(* IEC 61131-3 sources: daoli-st-library/DL_Process (part 58) *)

(* ---- FB_DL_VacuumBakeOutSeq.st ---- *)
(*
  组件名 Component   : FB_DL_VacuumBakeOutSeq
  子库 Sublibrary    : DL_Process
  版本 Version       : 1.0.0
  兼容性 Platform    : CODESYS 3.5 / TwinCAT 3 / 汇川 InoProShop / Machine Expert（仅 Standard.library）
  功能 Function      : 真空烘烤顺控（锂电/半导体共性，自研行业池）：
                       1) 升温相（eRampUp）：温度需求按 fRampRateKMin 斜率逼近
                       fSoakTempC，腔压 < fSoakPressMaxPa 才视为升温有效；
                       2) 保温保压相（eSoak）：温度需求保持 fSoakTempC，腔压超上限
                       持续 tPressDevTo → 故障锁存；保温计时到 → 进压升率判漏相；
                       3) 压升率判漏相（eRorMeas）：窗始取腔压快照，窗长 tRorWin 到
                       → 压升率 = (腔压 - 快照) / 窗长，超 fRorFailPaS → 故障（判漏
                       不合格）；不超 → 终点判据达成，进降温相；
                       4) 降温放气相（eCoolVent）：需求温度按斜率降至 fEndTempC 后
                       开放气阀驻留 tVentDur → eDone。
  边界 Boundary      : ① 本件只出温度需求/阀门指令，不写物理 IO，不内嵌温控回路；
                       ② 压升率除法前置域闸：tRorWin 秒值下限 0.1 s（常量护栏）；
                       ③ 各相计时独立 TON 实例（禁跨相复用）；压升率窗始快照在
                       进相首拍写定，锁存回放不重扫；
                       ④ 故障锁存解除唯一路径 = bReset 上升沿（输入引脚，恒可达）；
                       ⑤ 无全局变量引用、无外部变量声明、无物理地址寻址。
  依赖 Depends       : Standard.library（R_TRIG / TON）
  溯源 Origin        : 道莅自研 clean-room（自研行业池：锂电/半导体真空烘烤共性
                       语义，零外部代码行复制）
  码位 Code          : 16#06_0_BF（Process 段 0006，B 子带 BF 格）
  码表 Error codes（本件格 06_0_BF，单轨子道：故障 0x02BF / 信息 0x01BF）:
    16#0006_02BF 故障级：烘烤顺控故障总码（保压越限 / 压升率判漏不合格 /
                 组态非法 / 输入非有限），锁存至复位
    16#0006_01BF 信息级：压升率判漏通过沿（进降温相迁移拍）
  修订历史 Revision  :
    2026-11-19  v1.0.0  R44 首版（批次 4 · 序号 16）
*)

TYPE E_DL_VboPhase :
(
    eIdle     := 0,   // 空闲：未使能 / Idle, not enabled
    eRampUp   := 10,  // 升温：斜坡逼近保温温度 / Ramping to soak temperature
    eSoak     := 20,  // 保温保压：保持温度与压力 / Soaking temperature and pressure
    eRorMeas  := 30,  // 判漏：压升率测量窗 / Rate-of-rise measurement window
    eCoolVent := 40,  // 降温放气：斜坡降温 + 放气 / Cooling and venting
    eDone     := 50,  // 完成：终点驻留 / Done, endpoint held
    eFault    := 90   // 故障：总码锁存 / Fault, latched
);
END_TYPE

FUNCTION_BLOCK FB_DL_VacuumBakeOutSeq
VAR_INPUT
    bEnable      : BOOL;                   // 使能（电平）[-] / Enable
    bReset       : BOOL;                   // 上升沿清故障锁存 [-] / Reset edge
    fChamberTempC: REAL;                   // 腔体实测温度 [摄氏度] / Chamber temperature
    fChamberPressPa: REAL;                 // 腔体实测压力 [帕斯卡] / Chamber pressure
    fSoakTempC   : REAL := 80.0;           // 保温温度 [摄氏度] / Soak temperature
    fEndTempC    : REAL := 35.0;           // 降温终点温度 [摄氏度] / Cool-down end temperature
    fRampRateKMin: REAL := 2.0;            // 升降温斜率 [开尔文/分] / Ramp rate
    fSoakPressMaxPa: REAL := 50.0;         // 保温压力上限 [帕斯卡] / Soak pressure ceiling
    fRorFailPaS  : REAL := 5.0;            // 压升率判漏限 [帕/秒] / Rate-of-rise fail limit
    tSoakDur     : TIME := T#24H;          // 保温时长 [毫秒] / Soak duration
    tRorWin      : TIME := T#60S;          // 压升率测量窗 [毫秒] / ROR measurement window
    tPressDevTo  : TIME := T#30S;          // 保压越限确认窗 [毫秒] / Pressure deviation timeout
    tVentDur     : TIME := T#60S;          // 放气驻留 [毫秒] / Vent dwell
    tCycle       : TIME := T#1S;           // 扫描周期 [毫秒] / Scan cycle time
END_VAR
VAR_OUTPUT
    fTempDemandC : REAL;                   // 温度需求输出 [摄氏度] / Temperature demand
    bPumpCmd     : BOOL;                   // 抽真空维持指令（升温/保温/判漏相）[-] / Vacuum maintain command
    bVentCmd     : BOOL;                   // 放气阀指令（放气驻留相电平）[-] / Vent valve command
    fRorPaS      : REAL;                   // 实测压升率 [帕/秒] / Measured rate of rise
    ePhase       : E_DL_VboPhase;          // 相位出口，段尾单点映射 / Phase outlet
    bError       : BOOL;                   // 故障锁存标志 [-] / Fault latch flag
    uErrId       : UDINT;                  // 事件码，0 = 无事件 / Event code
END_VAR
VAR
    rtReset  : R_TRIG;                     // 复位沿实例，段 0 无条件刷新 / Reset edge
    tonSoakDur: TON;                       // 保温计时（独立实例） / Soak duration timer
    tonRorWin : TON;                       // 压升率测量窗（独立实例） / ROR window timer
    tonPressDevTo: TON;                    // 保压越限确认（专用超时件命名） / Pressure timeout
    tonVentDur: TON;                       // 放气驻留计时（独立实例） / Vent dwell timer
    _ePhase : E_DL_VboPhase := E_DL_VboPhase.eIdle;    // 内部相位（CASE 唯一写入目标）/ Internal phase
    _fPressSnap: REAL;                     // 判漏窗始压力快照 [帕斯卡] / Window-start pressure snapshot
    _fPressStart: REAL;                    // 保温起点压力快照 [帕斯卡] / Soak-start pressure snapshot
    _bFault : BOOL;                        // 故障锁存位（锁存量） / Latched fault bit
    _uFault : UDINT;                       // 故障码锁存（锁存量） / Latched fault code
    _bCfgBad: BOOL;                        // 组态非法当拍量 [-] / Config illegal flag
    _bNonFin: BOOL;                        // 输入非有限当拍量 [-] / Non-finite input flag
    _bSnapDone: BOOL;                      // 判漏快照已取标志 [-] / Snapshot taken flag
END_VAR
VAR CONSTANT
    DL_WIN_MIN_S : REAL := 0.1;            // 测量窗秒值下限 [秒] / Window seconds floor
    DL_SEC_PER_MIN: REAL := 60.0;          // 秒 → 分换算系数 [秒/分] / Seconds per minute
    DL_MS_PER_S  : REAL := 1000.0;         // 毫秒 → 秒换算系数 [毫秒/秒] / Milliseconds per second
    DL_ABS_MAX   : REAL := 1.0E30;         // 有限值判定上界 [工程单位] / Finite bound
    DL_ZERO      : REAL := 0.0;            // 零常量 [工程单位] / Zero constant
END_VAR

(* —— 段 0｜沿与定时器每拍无条件刷新（禁置于 IF/CASE 内；各相独立实例禁复用） —— *)
rtReset(CLK := bReset);
tonSoakDur   (IN := (_ePhase = E_DL_VboPhase.eSoak) AND (NOT _bFault), PT := tSoakDur);
tonRorWin    (IN := (_ePhase = E_DL_VboPhase.eRorMeas) AND (NOT _bFault), PT := tRorWin);
tonPressDevTo(IN := (_ePhase = E_DL_VboPhase.eSoak) AND (fChamberPressPa > fSoakPressMaxPa)
              AND (NOT _bFault), PT := tPressDevTo);
tonVentDur   (IN := (_ePhase = E_DL_VboPhase.eCoolVent) AND (NOT _bFault), PT := tVentDur);

(* —— 段 1｜瞬时量预清零（锁存量 _bFault/_uFault/fTempDemandC/_fPressSnap 不入清单） —— *)
uErrId   := 16#0000_0000;
_bCfgBad := FALSE;
_bNonFin := FALSE;

(* —— 段 2｜复位沿：故障一次性清干净，相位回空闲，阀门指令撤销 —— *)
IF rtReset.Q THEN
    _bFault := FALSE;
    _uFault := 16#0000_0000;
    bVentCmd := FALSE;
    bPumpCmd := FALSE;
    _ePhase := E_DL_VboPhase.eIdle;
END_IF

(* —— 段 3｜组态闸与非有限判据（覆盖全部参与判据换算引脚） —— *)
IF (fRampRateKMin <= DL_ZERO) OR (fRorFailPaS <= DL_ZERO) OR (tSoakDur = T#0S)
   OR (tRorWin = T#0S) OR (tPressDevTo = T#0S) OR (tVentDur = T#0S) OR (tCycle = T#0S)
   OR (fSoakTempC <= fEndTempC) THEN
    _bCfgBad := TRUE;
END_IF
IF (fChamberTempC <> fChamberTempC) OR ((fChamberTempC - fChamberTempC) <> DL_ZERO)
   OR (fChamberPressPa <> fChamberPressPa) OR ((fChamberPressPa - fChamberPressPa) <> DL_ZERO) THEN
    _bNonFin := TRUE;
END_IF

(* —— 段 4｜主状态机：七态全覆盖 + ELSE 兜底 —— *)
CASE _ePhase OF

E_DL_VboPhase.eIdle:
    fTempDemandC := fChamberTempC;       // 空闲相：需求跟随实测（不驱动）
    bPumpCmd := FALSE;
    bVentCmd := FALSE;
    IF bEnable AND (NOT _bCfgBad) THEN
        _bSnapDone := FALSE;
        fRorPaS := DL_ZERO;
        _ePhase := E_DL_VboPhase.eRampUp;
    ELSIF bEnable AND _bCfgBad THEN
        _bFault := TRUE;
        _uFault := 16#0006_02BF;
        bError  := TRUE;
        _ePhase := E_DL_VboPhase.eFault;
    END_IF

E_DL_VboPhase.eRampUp:
    bPumpCmd := TRUE;
    bVentCmd := FALSE;
    (* 温度需求斜率逼近：每拍步长 = 斜率 × 周期（分 → 秒换算，除子域闸已过） *)
    fTempDemandC := MIN(fTempDemandC + fRampRateKMin * (TIME_TO_REAL(tCycle) / DL_MS_PER_S)
                        / DL_SEC_PER_MIN, fSoakTempC);
    IF _bNonFin THEN
        _bFault := TRUE;
        _uFault := 16#0006_02BF;
        bError  := TRUE;
        _ePhase := E_DL_VboPhase.eFault;
    ELSIF NOT bEnable THEN
        _ePhase := E_DL_VboPhase.eIdle;  // 使能撤销回空闲
    ELSIF (fChamberTempC >= fSoakTempC) AND (fChamberPressPa <= fSoakPressMaxPa) THEN
        _fPressStart := fChamberPressPa; // 保温起点压力快照
        _ePhase := E_DL_VboPhase.eSoak;  // 迁出：温度达保温且压力已入保压域
    END_IF

E_DL_VboPhase.eSoak:
    bPumpCmd := TRUE;
    bVentCmd := FALSE;
    fTempDemandC := fSoakTempC;          // 保温相需求定值
    IF _bNonFin OR tonPressDevTo.Q THEN
        _bFault := TRUE;                 // 保压越限或输入非法：锁存
        _uFault := 16#0006_02BF;
        bError  := TRUE;
        _ePhase := E_DL_VboPhase.eFault;
    ELSIF NOT bEnable THEN
        _ePhase := E_DL_VboPhase.eIdle;  // 使能撤销回空闲
    ELSIF tonSoakDur.Q THEN
        _bSnapDone := FALSE;             // 保温时长到：进判漏相，快照待取
        _ePhase := E_DL_VboPhase.eRorMeas;
    END_IF

E_DL_VboPhase.eRorMeas:
    bPumpCmd := TRUE;
    bVentCmd := FALSE;
    fTempDemandC := fSoakTempC;
    IF _bNonFin THEN
        _bFault := TRUE;
        _uFault := 16#0006_02BF;
        bError  := TRUE;
        _ePhase := E_DL_VboPhase.eFault;
    ELSIF NOT _bSnapDone THEN
        _fPressSnap := fChamberPressPa;  // 窗始快照：进相首拍写定（锁存回放不重扫）
        _bSnapDone := TRUE;
    ELSIF tonRorWin.Q THEN
        (* 压升率 = (腔压 - 窗始快照) / 窗长秒值（除子 = 窗长，常量护栏下限已过） *)
        fRorPaS := (fChamberPressPa - _fPressSnap)
                   / MAX(TIME_TO_REAL(tRorWin) / DL_MS_PER_S, DL_WIN_MIN_S);
        IF fRorPaS > fRorFailPaS THEN
            _bFault := TRUE;             // 判漏不合格：锁存（禁按当下输入重推断）
            _uFault := 16#0006_02BF;
            bError  := TRUE;
            _ePhase := E_DL_VboPhase.eFault;
        ELSE
            uErrId := 16#0006_01BF;      // 信息级：判漏通过沿
            _ePhase := E_DL_VboPhase.eCoolVent;   // 终点判据达成：进降温放气
        END_IF
    END_IF

E_DL_VboPhase.eCoolVent:
    bPumpCmd := FALSE;
    (* 温度需求斜率下降，降至终点温度前放气阀不开（先降温后放气） *)
    IF fTempDemandC > fEndTempC THEN
        fTempDemandC := MAX(fTempDemandC - fRampRateKMin * (TIME_TO_REAL(tCycle) / DL_MS_PER_S)
                            / DL_SEC_PER_MIN, fEndTempC);
        bVentCmd := FALSE;
    ELSE
        bVentCmd := TRUE;                // 需求到终点温度：开放气阀驻留
    END_IF
    IF _bNonFin THEN
        _bFault := TRUE;
        _uFault := 16#0006_02BF;
        bError  := TRUE;
        _ePhase := E_DL_VboPhase.eFault;
    ELSIF bVentCmd AND tonVentDur.Q THEN
        _ePhase := E_DL_VboPhase.eDone;  // 迁出：放气驻留完成
    ELSIF NOT bEnable THEN
        _ePhase := E_DL_VboPhase.eIdle;  // 使能撤销回空闲
    END_IF

E_DL_VboPhase.eDone:
    bPumpCmd := FALSE;
    bVentCmd := FALSE;                   // 完成相：阀门指令全撤（安全侧）
    IF NOT bEnable THEN
        _ePhase := E_DL_VboPhase.eIdle;  // 使能撤销回空闲（待机可返回路径）
    END_IF

E_DL_VboPhase.eFault:
    bPumpCmd := FALSE;
    bVentCmd := FALSE;
    bError := TRUE;
    ;                                    // 故障相驻留：只认复位沿（段 2 迁出）

ELSE
    _bFault := TRUE;                     // 兜底：非法相位锁存
    _uFault := 16#0006_02BF;
    bError  := TRUE;
    _ePhase := E_DL_VboPhase.eFault;
END_CASE

(* —— 段 5｜相位出口单点映射 —— *)
ePhase := _ePhase;
END_FUNCTION_BLOCK

(* ---- FB_DL_VacuumChamberSeq.st ---- *)
(*==============================================================================
 * 组件名称 (Component)  : FB_DL_VacuumChamberSeq
 * 所属子库 (Sublibrary) : DL_Process
 * 前缀     (Prefix)     : FB_DL_
 * 当前版本 (Version)    : 1.0.0
 * 兼容性   (Platform)   : CODESYS 3.5 / TwinCAT 3 / 汇川 InoProShop / Schneider
 *                         Machine Expert；纯 IEC 61131-3（第 3 版），
 *                         仅依赖标准库 TON / R_TRIG / ABS，零厂商方言
 * 作者     (Author)     : 道莅代码库 · PLC编程专家（R31）
 * 开源溯源 (Origin)     : 真空腔体抽真空顺控公开工艺语义（行业池），
 *                         道莅 clean-room 防御性实现，未复制任何外部源码行
 * 功能描述 (Function)   : 纯真空腔体五相顺控原子（不含工艺加热）：粗抽至
 *                         粗抽阈值 → 精抽至目标（迟滞防边界抖动）→ 检漏
 *                         （消费 bLeakOk）→ 放气（数字阀经缓启时序等价
 *                         斜坡限幅防冲击）→ 完成。相转换本拍复验数据源
 *                         （R42）；步超时锁故障；中止安全次序写死：
 *                         先停泵、延时后才开放气阀。
 * 组合建议 (Composition): 与库内 FB_DL_SlitValveInterlock 组合使用——本件
 *                         给出真空工艺时序，闸阀联锁由该件承担，二者经
 *                         bLeakOk/泵指令引脚对接，不互相内嵌。
 * 状态机   (States)     : eIdle/eRough/eFine/eLeakTest/eVent/eFault，
 *                         CASE 带 ELSE 锁安全侧（全阀关、全泵停）。
 * 码位     (Codes)      : 16#0005_009E 信息级：压强数据非有限冻结当前相、
 *                                      迟滞等待提示（不置 bError）
 *                         16#0005_009F 故障级：相超时
 *                         16#0005_00A0 故障级：联锁违例（非空闲相重启）
 *                         16#0005_00A1 故障级：状态非法（ELSE 兜底，锁存）
 *                         16#0005_00A2 保留未启用（码表与实现对齐）
 * 边界防错 (Boundary)   : 1 压强非有限（x<>x 自反判加幅值界）冻结当前相；
 *                         2 精抽到位判定带迟滞：超回差即回信息级等待；
 *                         3 TON/R_TRIG 实例每拍无条件刷新，按相断输入；
 *                         4 CASE 带 ELSE 锁安全侧；
 *                         5 故障锁存可达解除路径：中止沿复归待机；
 *                         6 相转换本拍复验数据源（R42）。
 * 修订历史 (Revision)   : 2026-11-18 v1.0.0 首版入库（R31 · 阶段三 · 序 12）
 *==============================================================================*)

(*------------------------------------------------------------------------------
 * 枚举: E_DL_VacPhase（归属本功能块，同文件发布，全库唯一属主）
 *----------------------------------------------------------------------------*)
TYPE E_DL_VacPhase :
(
    eIdle     := 0,    // 空闲：全泵停全阀关 / Idle, all pumps and valves off
    eRough    := 10,   // 粗抽相：粗抽泵运行 / Rough phase, rough pump running
    eFine     := 20,   // 精抽相：精抽泵运行 / Fine phase, fine pump running
    eLeakTest := 30,   // 检漏相：泵停隔离等待结论 / Leak test, pumps off, isolated
    eVent     := 40,   // 放气相：缓启时序后开阀 / Vent phase, valve after ramp delay
    eFault    := 99    // 故障：锁定等待中止复位 / Fault, latched until abort reset
);
END_TYPE

(*==============================================================================
 * 功能块: FB_DL_VacuumChamberSeq
 * 调用约定: 每个扫描周期无条件调用一次；压强信号经引脚注入。
 *==============================================================================*)
FUNCTION_BLOCK FB_DL_VacuumChamberSeq
VAR_INPUT
    bStart   : BOOL := FALSE;         // 启动沿（空闲相受理）/ Start edge, accepted in idle
    bAbort   : BOOL := FALSE;         // 中止沿：任意相安全退出 / Abort edge, safe exit from any phase
    fPNow    : REAL := 101325.0;      // 腔体当前压强 [帕] / Chamber current pressure [Pa]
    fPTgt    : REAL := 10.0;          // 精抽目标压强 [帕] / Fine target pressure [Pa]
    fPRough  : REAL := 500.0;         // 粗抽切换阈值 [帕] / Rough crossover threshold [Pa]
    bLeakOk  : BOOL := FALSE;         // 检漏结论注入（外部检漏件）/ Leak verdict injected by caller
    tStepMax : TIME := T#600S;        // 单相超时 [毫秒] / Per-phase timeout [ms]
    tVentRamp: TIME := T#5S;          // 放气缓启时序 [毫秒]（斜坡限幅等价实现）/ Vent ramp delay [ms]
END_VAR
VAR_OUTPUT
    ePhase    : E_DL_VacPhase;        // 当前相状态 / Current phase
    bPumpRough: BOOL;                 // 粗抽泵指令 / Rough pump command
    bPumpFine : BOOL;                 // 精抽泵指令 / Fine pump command
    bVent     : BOOL;                 // 放气阀指令 / Vent valve command
    bDone     : BOOL;                 // 流程完成单拍脉冲（R27）/ Sequence done one-scan pulse
    bError    : BOOL;                 // 故障标志，与故障级码配对（R45）/ Fault flag paired with fault codes
    uErrorId  : UDINT;                // 错误码，0 = 无错 / Error code, 0 = none
END_VAR
VAR
    rTrigStart: R_TRIG;               // 启动沿检测，每拍无条件刷新 / Start edge detector, refreshed every scan
    rTrigAbort: R_TRIG;               // 中止沿检测，每拍无条件刷新 / Abort edge detector, refreshed every scan
    tonPhase  : TON;                  // 相超时定时器，每拍无条件刷新 / Phase timeout timer, refreshed every scan
    tonVent   : TON;                  // 放气缓启定时器，每拍无条件刷新 / Vent ramp timer, refreshed every scan
    eStatePrev: E_DL_VacPhase;        // 上一拍相快照 / Previous phase snapshot
    bStepRst  : BOOL;                 // 相切换拍单拍断超时输入 / One-scan timeout break on phase change
    bDataOk   : BOOL;                 // 压强三点有效性 / Three pressure points validity
    bHystWait : BOOL;                 // 迟滞等待标志 / Hysteresis waiting flag
    bAborted  : BOOL;                 // 中止退出路径标志 / Abort exit path flag
    uCodeLatch: UDINT;                // 故障级锁存码 / Latched fault code
    bInit     : BOOL := TRUE;         // 首扫标志 / First-scan flag
END_VAR
VAR CONSTANT
    DL_VCS_FIN    : REAL := 1.0E30;   // REAL 有限幅值判界 / REAL finiteness magnitude bound
    DL_VCS_HYST   : REAL := 1.1;      // 精抽迟滞回差系数（超回差回等待）/ Fine hysteresis back factor
    DL_VCS_PATM   : REAL := 90000.0;  // 放气完成压强阈 [帕] / Vent complete pressure threshold [Pa]
END_VAR

// ---- 段 1｜边沿与定时器实例无条件周期刷新（红线：禁入条件分支）----------------
rTrigStart(CLK := bStart);                            // 启动沿检测 / Start edge detection
rTrigAbort(CLK := bAbort);                            // 中止沿检测 / Abort edge detection
tonVent(IN := (ePhase = eVent), PT := tVentRamp);     // 缓启计时按相断输入 / Ramp timing input per phase
tonPhase(IN := (ePhase <> eIdle) AND (ePhase <> eFault) AND (ePhase <> eVent)
         AND (NOT bStepRst), PT := tStepMax);         // 相超时计时，相切换拍断输入 / Phase timeout timing

// ---- 段 2｜相切换检测与数据有效性 ----------------------------------------------
bStepRst := (ePhase <> eStatePrev) OR bInit;          // 相变化即断输入 / Phase change breaks timing input
eStatePrev := ePhase;                                 // 快照留痕 / Snapshot previous phase
bInit := FALSE;                                       // 清首扫标志 / Clear first-scan flag
bDataOk := (fPNow = fPNow) AND (fPTgt = fPTgt) AND (fPRough = fPRough)
       AND (ABS(fPNow) < DL_VCS_FIN) AND (ABS(fPTgt) < DL_VCS_FIN)
       AND (ABS(fPRough) < DL_VCS_FIN);               // 压强三点有限 / Three points finite

// ---- 段 3｜中止沿统一入口：先停泵、缓启延时后才放气（安全次序写死）--------------
IF rTrigAbort.Q AND (ePhase <> eIdle) THEN
    ePhase   := eVent;                                // 转放气相执行退出 / To vent phase for exit
    bAborted := TRUE;                                 // 登记中止路径 / Mark abort path
END_IF

// ---- 段 4｜状态机（CASE 带 ELSE 锁安全侧：全泵停全阀关）--------------------------
CASE ePhase OF
    eIdle:
        bPumpRough := FALSE;                          // 空闲全停 / All off in idle
        bPumpFine  := FALSE;                          // 空闲全停 / All off in idle
        bVent      := FALSE;                          // 空闲阀关 / Valve closed in idle
        bDone      := FALSE;                          // 清完成脉冲 / Clear done pulse
        bAborted   := FALSE;                          // 清中止标志 / Clear abort flag
        IF rTrigStart.Q AND bDataOk AND (fPTgt < fPRough) THEN
            ePhase := eRough;                         // 数据合法且目标低于切换阈才启动 / Legal data and sane targets
        END_IF
    eRough:
        bPumpRough := bDataOk AND NOT bAborted;       // 粗抽泵指令带数据门控 / Rough pump gated by data
        bPumpFine  := FALSE;                          // 精抽泵停 / Fine pump off
        bVent      := FALSE;                          // 阀关 / Valve closed
        IF NOT bDataOk THEN
            uErrorId := 16#0005_009E;                 // 信息级：数据非有限冻结当前相 / Info: non-finite freezes phase
        ELSIF tonPhase.Q THEN
            ePhase := eFault;                         // 相超时锁故障 / Phase timeout, fault
            uCodeLatch := 16#0005_009F;               // 码位：相超时 / Code: phase timeout
        ELSIF bDataOk AND (fPNow <= fPRough) THEN
            ePhase := eFine;                          // 复验后转精抽（R42）/ Recheck then to fine
        END_IF
    eFine:
        bPumpRough := FALSE;                          // 粗抽泵停（交叉点切换）/ Rough pump off at crossover
        bPumpFine  := bDataOk AND NOT bAborted;       // 精抽泵指令带数据门控 / Fine pump gated by data
        bVent      := FALSE;                          // 阀关 / Valve closed
        bHystWait  := bDataOk AND (fPNow > fPTgt * DL_VCS_HYST); // 超回差等待 / Beyond hysteresis, wait
        IF NOT bDataOk THEN
            uErrorId := 16#0005_009E;                 // 信息级：数据非有限冻结当前相 / Info: non-finite freezes phase
        ELSIF tonPhase.Q THEN
            ePhase := eFault;                         // 相超时锁故障 / Phase timeout, fault
            uCodeLatch := 16#0005_009F;               // 码位：相超时 / Code: phase timeout
        ELSIF bHystWait THEN
            uErrorId := 16#0005_009E;                 // 信息级：迟滞等待提示 / Info: hysteresis waiting
        ELSIF bDataOk AND (fPNow <= fPTgt) THEN
            ePhase := eLeakTest;                      // 复验后转检漏（R42）/ Recheck then to leak test
        END_IF
    eLeakTest:
        bPumpRough := FALSE;                          // 检漏隔离全泵停 / Isolated, all pumps off
        bPumpFine  := FALSE;                          // 检漏隔离全泵停 / Isolated, all pumps off
        bVent      := FALSE;                          // 阀关 / Valve closed
        IF tonPhase.Q THEN
            ePhase := eFault;                         // 相超时锁故障 / Phase timeout, fault
            uCodeLatch := 16#0005_009F;               // 码位：相超时 / Code: phase timeout
        ELSIF bLeakOk THEN
            ePhase := eVent;                          // 检漏合格转放气 / Leak OK, to vent
        END_IF
    eVent:
        bPumpRough := FALSE;                          // 放气相全泵停 / All pumps off in vent
        bPumpFine  := FALSE;                          // 放气相全泵停 / All pumps off in vent
        bVent      := tonVent.Q;                      // 缓启时序满才开阀（先停泵后放气）/ Valve after ramp, pumps first
        IF (NOT bAborted) AND bDataOk AND (fPNow >= DL_VCS_PATM) THEN
            ePhase := eIdle;                          // 正常放气完成回待机 / Normal vent complete
            bDone := TRUE;                            // 完成单拍脉冲 / One-scan done pulse
        ELSIF bAborted AND tonVent.Q THEN
            ePhase := eIdle;                          // 中止退出回待机 / Abort exit back to idle
            bDone := FALSE;                           // 中止不置完成 / Abort never sets done
        END_IF
    eFault:
        bPumpRough := FALSE;                          // 故障安全侧全停 / Fault safe side all off
        bPumpFine  := FALSE;                          // 故障安全侧全停 / Fault safe side all off
        bVent      := FALSE;                          // 故障安全侧阀关 / Fault safe side valve closed
        bDone      := FALSE;                          // 故障清完成 / Fault clears done
        IF rTrigAbort.Q THEN
            ePhase := eIdle;                          // 可达解除路径：中止沿复归 / Reachable release: abort edge
            uCodeLatch := 16#0000_0000;               // 清锁存码 / Clear latched code
        END_IF
    ELSE
        ePhase := eFault;                             // 非法状态兜底 / Illegal state fallback
        uCodeLatch := 16#0005_00A1;                   // 码位：状态非法 / Code: illegal state
END_CASE

// ---- 段 5｜联锁违例防御：非空闲相受理启动沿 --------------------------------------
IF rTrigStart.Q AND (eStatePrev <> eIdle) AND (ePhase <> eIdle) AND (ePhase <> eFault) THEN
    ePhase := eFault;                                 // 违例锁故障 / Violation latches fault
    uCodeLatch := 16#0005_00A0;                       // 码位：联锁违例 / Code: interlock violation
END_IF

// ---- 段 6｜错误码装配：故障锁存回放优先，信息级居次 ------------------------------
IF ePhase = eFault THEN
    bError   := TRUE;                                 // 故障标志配对（R45）/ Fault flag paired
    uErrorId := uCodeLatch;                           // 故障码锁存回放 / Latched fault code replayed
ELSIF (NOT bDataOk) OR bHystWait THEN
    bError   := FALSE;                                // 信息级不置故障 / Info never sets fault
    uErrorId := 16#0005_009E;                         // 信息级：冻结/迟滞等待 / Info: frozen or hysteresis wait
ELSE
    bError   := FALSE;                                // 无错清标志 / Clear fault flag
    uErrorId := 16#0000_0000;                         // 无码 / No code
END_IF
END_FUNCTION_BLOCK

(* ---- FB_DL_VavCouplingFeedforward.st ---- *)
(*==============================================================================
 * 组件名称 (Component)  : FB_DL_VavCouplingFeedforward
 * 所属子库 (Sublibrary) : DL_Process
 * 归属目录 (Directory)  : C:\Library\DL_Process
 * 当前版本 (Version)    : 1.0.0
 * 分类/来源标签         : 功能块（FUNCTION_BLOCK）· 暖通前馈 · 变风量耦合
 *                         industry-pool / hvac / vav / feedforward
 * 兼容性   (Platform)   : CODESYS 3.5 / TwinCAT 3 / 汇川 InoProShop / 施耐德
 *                         Machine Expert；仅用 Standard.library 的 ABS
 * 溯源声明 (Provenance) : 道莅自研 clean-room——只借公开规范条款与工程惯例，零代码行复制。
 * 功能一句话 (Summary)  : 送风温度偏离设计值时按显热守恒比例前馈修正风量
 *                         给定，替代反馈环慢慢追赶，防送风温度-风量耦合振荡。
 *
 * 功能描述 (Function)   : 显热守恒：风量与（室温设定 − 送风温度）成反比，
 *                         前馈量 = 设计风量 × 设计温差 ÷ 当前温差；当前温差
 *                         绝对值小于容差时视为近设计工况，恒等输出设计风量
 *                         并报信息级；输入非有限冻结输出（故障级）；送风
 *                         过热（温差反号）按最小风量保守输出；结果钳位到
 *                         风量上下限并报钳位码。内部状态与输出模式分离，
 *                         输出预置不触碰状态驻留量（R19）。
 * 与既有件边界 (Boundary): 本件只做静态前馈，不含反馈环与执行器控制；
 *                         VAV 盒反馈控制归 FB_DL_VavBoxCtrl，二者级联使用。
 * 码位说明 (Codes)      : 信息 16#0006_300A 近设计工况恒等输出设计风量
 *                         故障 16#0006_300B 输入非有限，输出冻结
 *                         故障 16#0006_300C 送风过热（温差反号），按最小风量保守
 *                         故障 16#0006_300D 结果越限已钳位到风量上下限
 *                         段 16#06_0_0A~0E 首槽信息级、次槽起故障级。
 * 依赖说明 (Depends)    : 无 DL_ 内部依赖；仅 Standard.library 的 ABS。
 * 红线自检 (Redline)    : 零全局依赖 ｜ 零 VAR_EXTERNAL ｜ 零 %I/%Q ｜ 纯 IEC 标准库
 *                         除法前强制判零（温差容差闸）｜ 浮点比较带 fEps 容差
 *                         NaN/Inf 精确判据拦截 ｜ ENUM 配 CASE 且 ELSE 兜底
 *                         全变量双语同行注释 ｜ 无定时器实例
 * 修订历史 (Revision)   : 2026-11-18  v1.0.0  首版入库（R32 · 批 3）
 *============================================================================*)

FUNCTION_BLOCK FB_DL_VavCouplingFeedforward
VAR_INPUT
    bRun        : BOOL;                     // 前馈使能，假则输出设计风量并停算 / Enable, FALSE outputs the design flow
    fTsaC       : LREAL;                    // 送风温度 [degC] / Supply air temperature
    fTsaDesignC : LREAL := 13.0;            // 设计送风温度 [degC] / Design supply air temperature
    fRoomSetC   : LREAL := 24.0;            // 室温设定 [degC] / Room setpoint
    fQDesign    : LREAL := 500.0;           // 设计风量 [m3/h] / Design airflow
    fQMin       : LREAL := 100.0;           // 最小风量 [m3/h] / Minimum airflow
    fQMax       : LREAL := 1200.0;          // 最大风量 [m3/h] / Maximum airflow
    fDtEps      : LREAL := 0.5;             // 温差容差 [K]，低于此视为近设计 / Delta-T tolerance
    fEps        : LREAL := 1.0E-6;          // 浮点判零容差 [实数域] / Floating zero tolerance
END_VAR
VAR_OUTPUT
    eMode   : (eBypass := 0, eAuto := 1);       // 模式枚举输出：旁路/自动 / Mode output enum
    fQFf    : LREAL;                    // 前馈风量给定 [m3/h] / Feedforward airflow setpoint
    bClamp  : BOOL;                     // 钳位标志，结果被上下限裁剪时为真 / TRUE when the result was clamped
    bValid  : BOOL;                     // 前馈有效标志，冻结期间为假 / TRUE when the output is valid
    bError  : BOOL;                     // 故障标志，与故障码配对 / Fault flag paired with codes
    uErrorId: UDINT;                    // 事件码，0 表示无事件 / Event code, zero means none
END_VAR
VAR
    _eState   : (eStBypass := 0, eStAuto := 1);     // 内部状态机：旁路/自动，输出预置不触碰 / Internal state, never pre-set
    fDtDesign : LREAL;  // 设计温差 [K]，室温设定减设计送风温度 / Design delta-T
    fDtNow    : LREAL;  // 当前温差 [K] / Current delta-T
    fRatio    : LREAL;  // 温差比 [比值]，设计温差除当前温差 / Delta-T ratio
    fQCalc    : LREAL;  // 计算风量 [m3/h] / Calculated airflow
    bSigOk    : BOOL;   // 输入有效标志 / Input validity flag
    uCode     : UDINT;  // 码位暂存，出口单点写入 [码] / Code staging
END_VAR

(* 段 1｜输出预置（不触碰 _eState 状态驻留量，R19 预清零清单纪律）/ Pre-set outputs, the state stays resident *)
fQFf    := fQDesign;                // 默认输出设计风量 / Default output is the design flow
bClamp  := FALSE;
bValid  := FALSE;
bError  := FALSE;
uErrorId := 16#0000_0000;
uCode   := 16#0000_0000;
eMode   := eBypass;                 // 模式输出随内部状态在出口刷新 / Mode output refreshed at the exit

(* 段 2｜温差导出与输入有效性（NaN 自反、Inf 上限、风量域正）/ Delta-T and validity *)
fDtDesign := fRoomSetC - fTsaDesignC;   // 设计温差导出 / Design delta-T
fDtNow    := fRoomSetC - fTsaC;         // 当前温差导出 / Current delta-T
bSigOk := (fTsaC = fTsaC) AND (fQDesign = fQDesign)             // NaN 自反判据 / NaN reflexivity
          AND (ABS(fTsaC) < 1.0E308) AND (ABS(fQDesign) < 1.0E308)   // Inf 上限判据 / Inf limit
          AND (fQDesign > fEps) AND (fQMin > 0.0) AND (fQMax > fQMin);   // 风量域约束 / Flow domain

(* 段 3｜状态机主分派（ENUM 配 CASE，ELSE 兜底）/ State dispatch with ELSE interception *)
CASE _eState OF

    eStBypass:
        (* 本拍行为：旁路保持设计风量；使能且数据有效拍 N+1 进自动 / Hold design flow; arm when enabled *)
        IF bRun AND bSigOk THEN
            _eState := eStAuto;         // 拍 N 旁路相满足条件，拍 N+1 转自动 / To auto next scan
        END_IF

    eStAuto:
        (* 本拍行为：按显热守恒算前馈；撤使能回旁路，数据无效冻结输出 / Compute feedforward; freeze on bad data *)
        IF NOT bRun THEN
            _eState := eStBypass;       // 拍 N+1 回旁路 / Back to bypass next scan
            fQFf := fQDesign;           // 旁路输出设计风量 / Bypass outputs design flow
        ELSIF NOT bSigOk THEN
            fQFf := fQDesign;           // 冻结：保持设计风量，不发异常值 / Freeze at design flow
            bValid := FALSE;            // 有效标志撤 / Withdraw validity
            uCode := 16#0006_300B;      // 故障级：输入非有限 / Fault: non-finite input
        ELSIF fDtNow < -fDtEps THEN
            fQFf := fQMin;              // 送风过热：保守最小风量 / Overheated supply: conservative minimum
            bValid := TRUE;
            uCode := 16#0006_300C;      // 故障级：温差反号 / Fault: reversed delta-T
        ELSE
            IF ABS(fDtNow) < fDtEps THEN
                fQFf := fQDesign;       // 近设计工况：恒等输出 / Near design: identity output
                bValid := TRUE;
                uCode := 16#0006_300A;  // 信息级：近设计恒等 / Info: near-design identity
            ELSE
                (* 除零前置闸：温差已过容差闸，此处防御复检再除 / Defensive recheck before the division *)
                IF ABS(fDtNow) > fEps THEN
                    fRatio := fDtDesign / fDtNow;   // 温差比 / Delta-T ratio
                    fQCalc := fQDesign * fRatio;    // 前馈风量 / Feedforward flow
                    IF fQCalc < fQMin THEN
                        fQCalc := fQMin;            // 钳下限 / Clamp to minimum
                        bClamp := TRUE;
                    ELSIF fQCalc > fQMax THEN
                        fQCalc := fQMax;            // 钳上限 / Clamp to maximum
                        bClamp := TRUE;
                    END_IF
                    fQFf := fQCalc;     // 前馈输出 / Feedforward output
                    bValid := TRUE;
                    IF bClamp THEN
                        uCode := 16#0006_300D;      // 故障级：结果已钳位 / Fault: clamped
                    END_IF
                ELSE
                    fQFf := fQMax;      // 防御路：温差趋零按最大风量 / Defensive: max flow as delta-T vanishes
                    bValid := TRUE;
                    uCode := 16#0006_300D;
                END_IF
            END_IF
        END_IF

ELSE
    _eState := eStBypass;               // 非法状态拦截回旁路 / Illegal state to bypass
    fQFf := fQDesign;                   // 保守输出设计风量 / Conservative design flow
    uCode := 16#0006_300B;              // 故障级：状态越界 / Fault: state out of range
END_CASE

(* 段 4｜出口装配 / Exit assembly *)
eMode := eBypass;                       // 出口刷新模式输出 / Refresh the mode output at the exit
IF _eState = eStAuto THEN
    eMode := eAuto;                     // 自动相映射 / Auto mapping
END_IF
bError := (uCode >= 16#0006_300B) AND (uCode <= 16#0006_300D);  // 故障级码段判定 / Fault band check
uErrorId := uCode;                      // 码位单点写入 / Single write point
END_FUNCTION_BLOCK

(* ---- FB_DL_VavDischargeAirReset.st ---- *)
(*
  FB_DL_VavDischargeAirReset  —  送风温度重置（末端阀位加权平均 → 送风设定值） / VAV discharge-air reset from terminal damper weighted mean
  分类 Category : DL_Process
  版本 Version  : 1.0.0
  来源 Source   : t1-2-oscat — 末端重置族零检索深化
  溯源 Origin   : clean-room 实现，未复制任何源码行
  功能 Function : 1) 末端阀位有效性门控：权重 = 有效末端数量（阀位域 [0,100] 且有限），
                  加权平均 fWMean := SUM(有效阀位)/有效末端数；
                  2) 重置律：fAirSet := fBaseSet + fResetSpan × fWMean/100，输出钳位
                  [fSetMin, fSetMax]，钳位发生置信息级 0494；
                  3) 权重和 = 0（全部末端无效）→ 防除零退回默认设定值 fBaseSet +
                  信息级 0492（不置故障）；
                  4) 部分末端无效置信息级 0493；非有限阀位 → 036B 锁存；
                  质量判定 CASE 全覆盖 + ELSE 兜底落 036C。
  边界 Boundary : ① 组态闸：uTermCnt < 1 或 > 8、fResetSpan < 0、设定钳位域颠倒 → 036A；
                  ② 除零防御：有效末端数 >= 1 过闸后才做除法；
                  ③ 无 GVL 依赖：纯引脚输入输出，无外部变量引用，无物理 IO 地址。
  依赖 Depends  : 仅 Standard.library（ABS / LREAL 算术）
  码表 Error codes（Process 段 0005，窗口 036A~036C / 0492~0494）:
    16#0005_036A 故障级：组态非法（末端数界外 / 重置幅值为负 / 钳位域颠倒），锁存至 bReset
    16#0005_036B 故障级：阀位非有限（NaN 自反判），锁存至 bReset
    16#0005_036C 故障级：质量判定落 ELSE 兜底（非法质量 ID），锁存至 bReset
    16#0005_0492 信息级：全部末端无效，退回默认设定值
    16#0005_0493 信息级：部分末端无效提示（有效末端照常聚合）
    16#0005_0494 信息级：设定值钳位提示
  修订历史 Revision :
    2026-11-19  v1.0.0  R41 首版（批次 4 · 序号 4）
*)

TYPE E_DL_VarResetQual :
(
    eAllValid   := 0,    // 全部末端有效 / All terminals valid
    ePartValid  := 10,   // 部分末端无效 / Some terminals invalid
    eNoneValid  := 20    // 全部末端无效 / No terminal valid
);
END_TYPE

FUNCTION_BLOCK FB_DL_VavDischargeAirReset
VAR_INPUT
    aDamper      : ARRAY[1..8] OF LREAL;  // 末端阀位 [0..100 %] / Terminal damper positions
    uTermCnt     : UINT := 1;         // 末端数 [个]，域 1..8 / Terminal count
    fBaseSet     : LREAL := 18.0;     // 基础送风设定 [°C] / Base discharge-air setpoint
    fResetSpan   : LREAL := 2.0;      // 重置幅值 [K]，域 >= 0（阀位 100% 时加满）/ Reset span
    fSetMin      : LREAL := 12.0;     // 设定值下限 [°C] / Setpoint lower clamp
    fSetMax      : LREAL := 26.0;     // 设定值上限 [°C] / Setpoint upper clamp
    bEnable      : BOOL := FALSE;     // 使能 [-] / Enable
    bReset       : BOOL := FALSE;     // 复位，上升沿清故障锁存 / Reset edge clears fault latch
END_VAR
VAR_OUTPUT
    fAirSet      : LREAL;             // 送风设定值出口 [°C] / Discharge-air setpoint outlet
    fWMean       : LREAL;             // 阀位加权平均 [0..100 %] / Weighted damper mean
    bValid       : BOOL;              // 输出有效标志 / Output valid flag
    bError       : BOOL;              // 故障锁存标志 / Fault latch flag
    nErrId       : UDINT;             // 事件码，0 = 无事件 / Event code
END_VAR
VAR
    rtReset      : R_TRIG;            // 复位沿实例，无条件刷新 / Reset edge instance
    _nCap        : INT;               // 生效末端数 [个] / Effective terminal count
    _nValid      : INT;               // 有效末端数 [个] / Valid terminal count
    _fSum        : LREAL;             // 阀位累加器 [0..100 %] / Damper sum accumulator
    _eQual       : E_DL_VarResetQual; // 质量判定（CASE 唯一写入目标）/ Quality verdict
    _bFault      : BOOL;              // 故障锁存位（锁存量）/ Latched fault bit
    _uFault      : UDINT;             // 故障码锁存（锁存量）/ Latched fault code
    _uInfo       : UDINT;             // 信息码，每拍重算 / Transient info code
    i            : INT;               // 聚合循环游标 [索引] / Aggregation loop cursor
    _nGuard      : INT;               // 聚合守卫计数 [次] / Aggregation guard counter
END_VAR

(* —— 段 0：沿实例无条件周期刷新（禁置于 IF/CASE 内） —— *)
rtReset(CLK := bReset);             // 复位沿（每拍必调）

(* —— 段 1：单拍量预清零（锁存量 _bFault/_uFault 不入清单，禁同拍抹除） —— *)
_uInfo := 16#0000_0000;             // 信息码每拍重算
bValid := FALSE;                    // 有效出口缺省 FALSE
nErrId := 16#0000_0000;             // 事件码缺省无事件
fAirSet := fBaseSet;                // 设定值缺省 = 默认设定值（退回口径）
fWMean := 0.0;                      // 均值缺省 0
_nValid := 0;                       // 有效计数清零
_fSum := 0.0;                       // 累加器清零
_nGuard := 0;                       // 守卫清零

(* —— 段 2：复位沿 + 组态域闸（当拍量判据） —— *)
IF rtReset.Q THEN                   // rtReset.Q = 当拍量
    _bFault := FALSE;               // 清故障锁存位
    _uFault := 16#0000_0000;        // 清故障锁存码
END_IF
_nCap := UINT_TO_INT(uTermCnt);     // 末端数快照
IF (_nCap < 1) OR (_nCap > 8) OR (fResetSpan < 0.0) OR (fSetMin >= fSetMax) THEN
    _uFault := 16#0005_036A;        // 故障级：组态非法
    _bFault := TRUE;
END_IF

(* —— 段 3：末端聚合（有效性门控；非有限 → 036B 锁存；守卫循环） —— *)
IF (NOT _bFault) AND (_nCap >= 1) AND (_nCap <= 8) THEN
    FOR i := 1 TO _nCap DO
        _nGuard := _nGuard + 1;     // 守卫递增
        IF _nGuard > 8 THEN
            EXIT;                   // 守卫兜底退出（理论不可达）
        END_IF
        IF (aDamper[i] <> aDamper[i]) OR ((aDamper[i] - aDamper[i]) <> (aDamper[i] - aDamper[i])) THEN
            _uFault := 16#0005_036B;    // 故障级：阀位非有限
            _bFault := TRUE;
        ELSIF (aDamper[i] >= 0.0) AND (aDamper[i] <= 100.0) THEN
            _nValid := _nValid + 1;     // 有效末端计数（权重 = 有效性门控）
            _fSum := _fSum + aDamper[i];    // 阀位累加
        END_IF
    END_FOR
END_IF

(* —— 段 4：质量判定（CASE 全覆盖 + ELSE 兜底） —— *)
IF (NOT _bFault) AND (_nCap >= 1) AND (_nCap <= 8) THEN
    IF _nValid = _nCap THEN
        _eQual := E_DL_VarResetQual.eAllValid;      // 全部有效
    ELSIF _nValid >= 1 THEN
        _eQual := E_DL_VarResetQual.ePartValid;     // 部分有效
        _uInfo := 16#0005_0493;                     // 信息级：部分无效提示
    ELSE
        _eQual := E_DL_VarResetQual.eNoneValid;     // 全部无效
    END_IF

    CASE _eQual OF
    E_DL_VarResetQual.eAllValid:
        fWMean := _fSum / INT_TO_LREAL(_nValid);    // 加权平均（分母 = 末端数 >= 1，防除零）
    E_DL_VarResetQual.ePartValid:
        fWMean := _fSum / INT_TO_LREAL(_nValid);    // 有效末端口径平均（同上防除零）
    E_DL_VarResetQual.eNoneValid:
        fWMean := 0.0;                              // 无有效样本
        _uInfo := 16#0005_0492;                     // 信息级：退回默认设定值
        fAirSet := fBaseSet;                        // 防除零退默认
    ELSE
        _uFault := 16#0005_036C;                    // 故障级：非法质量 ID 兜底
        _bFault := TRUE;
        fAirSet := fBaseSet;                        // 安全侧退默认
    END_CASE
END_IF

(* —— 段 5：重置律与钳位（分母 100.0 为常量恒非零） —— *)
IF (NOT _bFault) AND (_nValid >= 1) THEN
    fAirSet := fBaseSet + fResetSpan * fWMean / 100.0;  // 重置律
    IF fAirSet < fSetMin THEN
        fAirSet := fSetMin;         // 下界钳位
        _uInfo := 16#0005_0494;     // 信息级：钳位提示
    ELSIF fAirSet > fSetMax THEN
        fAirSet := fSetMax;         // 上界钳位
        _uInfo := 16#0005_0494;     // 信息级：钳位提示
    END_IF
END_IF

(* —— 段 6：出口单点映射（锁存码回放，禁同拍抹除） —— *)
bValid := (NOT _bFault) AND bEnable AND (_nValid >= 1);  // 有效出口
IF _bFault THEN
    nErrId := _uFault;              // 故障锁存码回放
    bValid := FALSE;                // 故障期强制 FALSE（安全侧）
    fAirSet := fBaseSet;            // 故障期退默认（安全侧）
ELSE
    nErrId := _uInfo;               // 信息码
END_IF
bError := _bFault;                  // 故障标志与锁存位同源

END_FUNCTION_BLOCK

(* ---- FB_DL_VffsBagLength.st ---- *)
(*==============================================================================
 * 组件名称 (Component)  : FB_DL_VffsBagLength
 * 所属子库 (Sublibrary) : DL_Process
 * 当前版本 (Version)    : 1.0.0
 * 兼容性 (Platform)     : CODESYS 3.5 / TwinCAT 3 / 汇川 InoProShop / Machine Expert
 *                         仅依赖纯 IEC 61131-3 标准元素，零厂商方言
 * 功能描述 (Function)   : 立式制袋袋长控制：编码器脉冲计长 → 色标上升沿比对基准
 *                         求偏差 → 偏差限幅后修正下一袋袋长；连续 N 袋（默认 3）
 *                         无色标 → bMarkLost 退化为定长（显式置位，不静默）；切刀
 *                         相位 = 计长对每袋脉冲取正余数，落对齐窗即就绪。
 *                         色标去抖 TON 5 ms 无条件刷新；模运算委托防负余数。
 * 溯源 (Origin)         : 道莅 clean-room 防御性实现
 * 本文件内含 (Contains) : TYPE E_DL_VffsErr / FUNCTION_BLOCK FB_DL_VffsBagLength
 * 依赖 (Depends)        : DL_MathData/FC_DL_ModPos
 * 红线自检 (Redline)    : 无外部全局变量、无硬件地址直引 ｜ 全变量中英双语同行注释
 *                         每袋脉冲为 0 拒绝（防除零）+ 修正双向钳制 + 模运算防负 ｜
 *                         枚举成员全部显式赋值 ｜ TON/R_TRIG 每周期无条件调用 ｜
 *                         退化态显式输出（不清零显示）｜ CASE 含 ELSE 兜底
 * 错误码表 (Codes)      : 16#0005_0417 同步运行
 *                         16#0005_0418 信息级 色标丢失（定长退化）
 *                         16#0005_0419 信息级 修正饱和（连续贴限）
 *                         16#0005_041A 故障级 编码器组态非法（每袋脉冲为 0）
 *                         16#0005_041B 信息级 相位对齐完成
 * 修订历史 (Revision)   : 2026-11-17  v1.0.0  首版入库 · R27 · 阶段三批 3
 * 验收向量 (Acceptance) : 每袋脉冲 1000、设定 300 mm：实测 1010 脉冲 → 偏差 +3 mm
 *                         → 下袋长 297 mm（限幅 5 mm 内）；连续 3 袋无标 → 0418 定长；
 *                         每袋脉冲 0 → 041A 拒绝
 *============================================================================*)

(*-----------------------------------------------------------------------------
 * 枚举: E_DL_VffsErr（归属 DL_Process，与 FB_DL_VffsBagLength 同文件）
 *----------------------------------------------------------------------------*)
TYPE E_DL_VffsErr :
(
    eSyncRun    := 16#0005_0417,   // 同步运行 / Synchronised running
    eMarkLost   := 16#0005_0418,   // 信息级：色标丢失，定长退化 / Info: mark lost, fixed-length degradation
    eCorrSat    := 16#0005_0419,   // 信息级：修正饱和（连续贴限）/ Info: correction saturated
    eEncBad     := 16#0005_041A,   // 故障级：编码器组态非法 / Fault: illegal encoder configuration
    ePhaseOk    := 16#0005_041B    // 信息级：相位对齐完成 / Info: cut phase aligned
);
END_TYPE

(*==============================================================================
 * 功能块: FB_DL_VffsBagLength
 * 调用约定: 每个扫描周期无条件调用一次；bEncPulse 必须注入真实编码器脉冲。
 *============================================================================*)
FUNCTION_BLOCK FB_DL_VffsBagLength
VAR_INPUT
    bMarkDetect   : BOOL;              // 色标传感器输入 / Mark sensor input
    bEncPulse     : BOOL;              // 编码器脉冲输入（计长源）/ Encoder pulse input, length source
    fBagLenSet_mm : REAL;              // 设定袋长 [毫米]，有效域 50~2000 / Set bag length [mm]
    uEncPpr       : UINT;              // 编码器每袋脉冲 [脉冲每袋]，须 > 0 / Encoder pulses per bag, must be > 0
    fCorrLimit_mm : REAL := 5.0;       // 修正限幅 [毫米]，默认 5 / Correction limit [mm]
    tMarkDeb      : TIME := T#5MS;     // 色标去抖时间 [毫秒]，默认 5 / Mark debounce time [ms]
    bReset        : BOOL;              // 复位（清丢失标记与修正）/ Reset, clears lost flag and correction
END_VAR
VAR_OUTPUT
    fBagLenAct_mm : REAL;              // 实际袋长（修正后，用于下一袋）[毫米] / Actual bag length, corrected [mm]
    fCorr_mm      : REAL;              // 当前修正量 [毫米] / Current correction [mm]
    bMarkLost     : BOOL;              // 色标丢失（定长退化）/ Mark lost, fixed-length degradation
    bCutPhaseOk   : BOOL;              // 切刀相位就绪 / Cut phase ready
    nEncCnt       : DINT;              // 当前袋内脉冲计数 [脉冲] / Pulse count in the current bag [pulses]
    nPhaseDiag    : DINT;              // 相位正余数诊断 [脉冲] / Positive-remainder phase diagnostic [pulses]
    eErr          : E_DL_VffsErr;      // 错误码 / Error code
END_VAR
VAR
    fbEncTrig     : R_TRIG;            // 编码器脉冲沿实例（无条件调用）/ Encoder pulse edge instance
    fbMarkTrig    : R_TRIG;            // 去抖后色标沿实例（无条件调用）/ Debounced mark edge instance
    fbResetTrig   : R_TRIG;            // 复位沿实例（无条件调用）/ Reset edge instance
    tonMarkDeb    : TON;               // 色标去抖定时器（无条件调用）/ Mark debounce timer
    fDev_mm       : REAL;              // 本袋脉冲偏差换算长度 [毫米] / Pulse deviation converted to length [mm]
    fCorrUse      : REAL;              // 修正量工作副本（钳位后）[毫米] / Correction working copy [mm]
    fPprUse       : REAL;              // 每袋脉冲实数副本（除子非零）[脉冲每袋] / Pulses per bag as real, non-zero
    uMissCnt      : UINT;              // 连续无色标袋数 [袋] / Consecutive bags without a mark [bags]
    uSatCnt       : UINT;              // 连续修正贴限次数 [次] / Consecutive saturated corrections [pcs]
    uPhaseWin     : DINT;              // 相位对齐窗宽 [脉冲] / Phase alignment window [pulses]
    uModErr       : UDINT;             // 委托取模错误码（0 = 无错）/ Delegate modulo error id
    bPprOk        : BOOL;              // 每袋脉冲合法性 / Pulses-per-bag legality
    bSatNow       : BOOL;              // 本袋修正贴限标志 / Correction saturated this bag
END_VAR
VAR CONSTANT
    DL_VFFS_LEN_MIN   : REAL := 50.0;    // 袋长域下限 [毫米] / Bag length lower bound [mm]
    DL_VFFS_LEN_MAX   : REAL := 2000.0;  // 袋长域上限 [毫米] / Bag length upper bound [mm]
    DL_VFFS_CORR_MIN  : REAL := 0.1;     // 修正限幅下限 [毫米] / Correction limit floor [mm]
    DL_VFFS_MISS_MAX  : UINT := 3;       // 连续无色标退化门限 [袋] / Mark-lost degradation threshold [bags]
    DL_VFFS_SAT_MAX   : UINT := 5;       // 连续贴限预警门限 [次] / Saturation warning threshold [pcs]
    DL_VFFS_WIN_DIV   : DINT := 20;      // 相位窗分数（每袋脉冲 / 20）/ Phase window divisor
    DL_VFFS_WIN_MIN   : DINT := 1;       // 相位窗最小宽 [脉冲] / Phase window minimum [pulses]
    DL_VFFS_MISS_FACT : DINT := 1;       // 无色标判据倍率（1 袋脉冲未到标即计一次丢标）/ Missing-mark pulse factor
    DL_VFFS_INF_MAX   : REAL := 1.0E30;  // 非有限值判定幅值上限 / Magnitude bound for finite-value check
    DL_VFFS_ZERO      : REAL := 0.0;     // 零值常量，避免裸字面量 / Zero constant
    DL_VFFS_EPS       : REAL := 0.001;   // 修正贴限比较容差 [毫米] / Saturation comparison tolerance [mm]
END_VAR

(*------------------------------------------------------------------------------
 * 段 1｜沿检测/TON 实例每周期无条件调用（仅输入条件化）
 *----------------------------------------------------------------------------*)
fbEncTrig(CLK := bEncPulse);                          // 编码器脉冲沿检测无条件刷新 / encoder edge refreshed unconditionally
tonMarkDeb(IN := bMarkDetect, PT := tMarkDeb);        // 色标去抖计时（无条件刷新）/ mark debounce timing
fbMarkTrig(CLK := tonMarkDeb.Q);                      // 去抖后色标沿检测无条件刷新 / debounced mark edge refreshed
fbResetTrig(CLK := bReset);                           // 复位沿检测无条件刷新 / reset edge refreshed

(*------------------------------------------------------------------------------
 * 段 2｜复位沿：清丢失标记、修正与计数
 *----------------------------------------------------------------------------*)
IF fbResetTrig.Q THEN
    bMarkLost := FALSE;                               // 丢失标记清 / lost flag cleared
    fCorrUse := DL_VFFS_ZERO;                         // 修正清 / correction cleared
    fCorr_mm := DL_VFFS_ZERO;                         // 修正输出清 / correction output cleared
    nEncCnt := 0;                                     // 计数清 / count cleared
    uMissCnt := 0;                                    // 丢标计数清 / miss count cleared
    uSatCnt := 0;                                     // 贴限计数清 / saturation count cleared
END_IF

(*------------------------------------------------------------------------------
 * 段 3｜编码器组态合法性与参数钳位（故障级 041A：每袋脉冲为 0 拒绝）
 *----------------------------------------------------------------------------*)
bPprOk := uEncPpr > 0;                                // 每袋脉冲合法判据 / pulses-per-bag legality
IF NOT bPprOk THEN
    eErr := E_DL_VffsErr.eEncBad;                     // 故障级：编码器组态非法 / fault: illegal encoder configuration
    bCutPhaseOk := FALSE;                             // 相位就绪撤（拒绝判定）/ phase ready dropped
    bMarkLost := TRUE;                                // 退化标记置位（显式，不清零显示）/ degradation flag explicit
    RETURN;
END_IF
IF (fBagLenSet_mm <> fBagLenSet_mm) OR (fBagLenSet_mm < DL_VFFS_LEN_MIN) OR (fBagLenSet_mm > DL_VFFS_LEN_MAX) THEN
    eErr := E_DL_VffsErr.eEncBad;                     // 袋长非法并入编码器组态段（反证句：同样拒绝判定）/ illegal length mapped to config band
    bCutPhaseOk := FALSE;                             // 相位就绪撤 / phase ready dropped
    RETURN;
END_IF
IF (fCorrLimit_mm <> fCorrLimit_mm) OR (fCorrLimit_mm < DL_VFFS_CORR_MIN) THEN
    fCorrLimit_mm := DL_VFFS_CORR_MIN;                // 修正限幅下限钳位（防除零式零限幅）/ correction limit floored
END_IF
fPprUse := UINT_TO_REAL(uEncPpr);                     // 每袋脉冲实数副本（非零已证）/ pulses per bag as real, proven non-zero

(*------------------------------------------------------------------------------
 * 段 4｜编码器计长：脉冲沿计数与本袋脉冲累计
 *----------------------------------------------------------------------------*)
IF fbEncTrig.Q THEN
    nEncCnt := nEncCnt + 1;                           // 本袋计数递增 [脉冲] / bag pulse count incremented
    IF nEncCnt > DL_VFFS_MISS_FACT * UINT_TO_DINT(uEncPpr) THEN
        nEncCnt := DL_VFFS_MISS_FACT * UINT_TO_DINT(uEncPpr);   // 计数上限钳位（防溢出与漂移累积）/ count capped
    END_IF
END_IF

(*------------------------------------------------------------------------------
 * 段 5｜色标沿：偏差换算、限幅、修正下一袋袋长，并清计数与丢标计数
 *----------------------------------------------------------------------------*)
eErr := E_DL_VffsErr.eSyncRun;                        // 默认码：同步运行 / default code: synchronised running
IF fbMarkTrig.Q THEN
    fDev_mm := (DINT_TO_REAL(nEncCnt) - fPprUse) / fPprUse * fBagLenSet_mm;   // 偏差换算 [毫米]（除子已证非零）/ deviation [mm]
    IF fDev_mm > fCorrLimit_mm THEN
        fDev_mm := fCorrLimit_mm;                     // 偏差上限钳制 / deviation capped
    ELSIF fDev_mm < -fCorrLimit_mm THEN
        fDev_mm := -fCorrLimit_mm;                    // 偏差下限钳制 / deviation floored
    END_IF
    fCorrUse := -fDev_mm;                             // 修正量取反（长袋则缩短下一袋）/ correction inverted for the next bag
    IF fCorrUse > fCorrLimit_mm THEN
        fCorrUse := fCorrLimit_mm;                    // 修正上限钳位 / correction capped
    ELSIF fCorrUse < -fCorrLimit_mm THEN
        fCorrUse := -fCorrLimit_mm;                   // 修正下限钳位 / correction floored
    END_IF
    bSatNow := ABS(fCorrUse) >= (fCorrLimit_mm - DL_VFFS_EPS);   // 本袋贴限判据（容差比较）/ saturated-this-bag predicate
    IF bSatNow THEN
        IF uSatCnt < DL_VFFS_SAT_MAX THEN
            uSatCnt := uSatCnt + 1;                   // 贴限计数递增 [次] / saturation count incremented
        END_IF
    ELSE
        uSatCnt := 0;                                 // 未贴限：贴限计数清零 / saturation count cleared
    END_IF
    fCorr_mm := fCorrUse;                             // 修正输出 [毫米] / correction output [mm]
    nEncCnt := 0;                                     // 本袋计数清零 / bag counter cleared
    uMissCnt := 0;                                    // 丢标计数清零 / miss count cleared
    bMarkLost := FALSE;                               // 色标恢复：退化解除 / mark recovered: degradation released
END_IF

(*------------------------------------------------------------------------------
 * 段 6｜色标丢失判定：计长超 2 袋仍未到标 → 丢标计数；连续 3 袋 → 定长退化
 *----------------------------------------------------------------------------*)
IF nEncCnt >= DL_VFFS_MISS_FACT * UINT_TO_DINT(uEncPpr) THEN
    IF uMissCnt < DL_VFFS_SAT_MAX THEN
        uMissCnt := uMissCnt + 1;                     // 丢标计数递增 [袋] / miss count incremented
    END_IF
    nEncCnt := 0;                                     // 计长清零（按定长循环计）/ counter cleared for fixed-length cycling
END_IF
IF uMissCnt >= DL_VFFS_MISS_MAX THEN
    bMarkLost := TRUE;                                // 连续丢标：定长退化（显式置位）/ mark lost: fixed-length degradation
    IF eErr = E_DL_VffsErr.eSyncRun THEN
        eErr := E_DL_VffsErr.eMarkLost;               // 信息级：色标丢失 / info: mark lost
    END_IF
END_IF
IF uSatCnt >= DL_VFFS_SAT_MAX THEN
    IF eErr = E_DL_VffsErr.eSyncRun THEN
        eErr := E_DL_VffsErr.eCorrSat;                // 信息级：修正饱和 / info: correction saturated
    END_IF
END_IF

(*------------------------------------------------------------------------------
 * 段 7｜袋长输出与切刀相位：模运算委托 FC_DL_ModPos 防负余数
 *----------------------------------------------------------------------------*)
fBagLenAct_mm := fBagLenSet_mm + fCorrUse;            // 实际袋长（修正后）[毫米] / actual bag length [mm]
IF fBagLenAct_mm < DL_VFFS_LEN_MIN THEN
    fBagLenAct_mm := DL_VFFS_LEN_MIN;                 // 袋长下限防护 / length floor
ELSIF fBagLenAct_mm > DL_VFFS_LEN_MAX THEN
    fBagLenAct_mm := DL_VFFS_LEN_MAX;                 // 袋长上限防护 / length ceiling
END_IF
nPhaseDiag := FC_DL_ModPos(nValue := nEncCnt, nModulus := UINT_TO_DINT(uEncPpr), eErr => uModErr);   // 相位正余数 [脉冲] / positive-remainder phase
IF uModErr <> 0 THEN
    nPhaseDiag := 0;                                  // 委托异常诊断归零 / diagnostic zeroed on delegate error
END_IF
uPhaseWin := UINT_TO_DINT(uEncPpr) / DL_VFFS_WIN_DIV;   // 相位窗宽 [脉冲] / phase window width [pulses]
IF uPhaseWin < DL_VFFS_WIN_MIN THEN
    uPhaseWin := DL_VFFS_WIN_MIN;                     // 窗宽下限钳位 / window floored
END_IF
bCutPhaseOk := (nPhaseDiag <= uPhaseWin) OR (nPhaseDiag >= (UINT_TO_DINT(uEncPpr) - uPhaseWin));   // 对齐窗判据 / alignment window predicate
IF bCutPhaseOk AND (eErr = E_DL_VffsErr.eSyncRun) THEN
    eErr := E_DL_VffsErr.ePhaseOk;                    // 信息级：相位对齐完成 / info: phase aligned
END_IF
END_FUNCTION_BLOCK

(* ---- FB_DL_VisionResultGate.st ---- *)
(*
  ==================================================================
  组件名 Component  : FB_DL_VisionResultGate
  分类   Category   : DL_Process
  复杂度 Complexity  : 中
  版本   Version    : 1.0.0
  功能   Purpose    : 视觉结果门控。工件到位沿开判决窗 tJudgeWin：窗内收到
                      结果选通（rtReady）按 bVisionOk 判 OK/NG；NG 可复检
                      （nRecheckMax 次上限）；窗超时无结果降级（bDegrade 单
                      脉冲 + nDegradeCnt 计数，安全侧判 NG 拒收）。TcOpen
                      视觉契约族范式，与 FB_DL_RobotGripVerify 分工。
  来源   Source     : T1-5-tcopen（TcOpen 视觉契约族范式）
  溯源   Origin     : 视觉判决窗与复检计数为公开工程范式，clean-room 自研
                      实现，未复制 TcOpen 或任何厂商私有库源码。
  平台   Platform   : 纯 IEC 61131-3（Standard.library: TON / R_TRIG，无私有库）
  分工声明 Split     : 与 FB_DL_RobotGripVerify 分工——后者做机器人抓取验
                      证，本件做视觉 OK/NG 判决门控。
  作者   Author     : 道莅代码库 · PLC 编程专家（R59）
  ------------------------------------------------------------------
  边界 Boundary     :
                      一 安全语义：降级（超时无结果）安全侧判 NG 拒收（R191
                         降级显式）；故障相输出全清；
                      二 判决窗到期即出（窗口末退出迁移，纪律④）；复检共用
                         同一窗口（迁相时窗续走不重启）；
                      三 bPass / bReject / bDegrade 均单拍脉冲，每拍前置清
                         零（纪律③防粘滞）；
                      四 组态域：nRecheckMax ∈ [0..9]，越域锁存 bError（解
                         除 = bReset 沿，R188）；
                      五 定时器与沿检测全部段 0 无条件周期刷新（R7）；
                      六 无全局变量、无外部变量声明、无物理地址寻址。
  修订记录 Revision  :
    2026-11-21  v1.0.0  R59 首版（批 4 · 序号 18）
  ==================================================================
*)

TYPE E_DL_VrgPhase :
(
    eVrgIdle    := 0,  // 空闲：等工件到位沿 / idle, awaiting the part edge
    eVrgJudge   := 10, // 判决窗：等结果选通 / the judge window, awaiting the result strobe
    eVrgRecheck := 20, // 复检窗：NG 后重判 / the recheck window after an NG
    eVrgFault   := 90  // 故障锁存：仅复位可清 / the latched fault
);
END_TYPE

FUNCTION_BLOCK FB_DL_VisionResultGate
VAR_INPUT
    bPartIn      : BOOL := FALSE; // 工件到位信号，上升沿开窗 [-] / the part in place signal, the rising edge opens the window
    bResultReady : BOOL := FALSE; // 视觉结果选通（结果有效单发）[-] / the result strobe, one shot valid
    bVisionOk    : BOOL := FALSE; // 视觉判决结果，TRUE = OK [-] / the vision verdict, true = ok
    tJudgeWin    : TIME := T#1S;  // 判决窗时长 [毫秒] / the judge window [millisecond]
    nRecheckMax  : INT  := 1;     // 复检次数上限 [次]，域 0..9 / the recheck bound, zero through nine
    bReset       : BOOL := FALSE; // 故障与组态复位，上升沿生效 [-] / the fault and config reset, rising edge
END_VAR
VAR_OUTPUT
    bPass        : BOOL := FALSE; // 判 OK 单脉冲（单拍）[-] / the pass one shot pulse, single scan
    bReject      : BOOL := FALSE; // 判 NG 拒收单脉冲（单拍）[-] / the reject one shot pulse, single scan
    bDegrade     : BOOL := FALSE; // 超时无结果降级单脉冲（单拍）[-] / the degrade one shot pulse, single scan
    nRecheckCnt  : INT  := 0;   // 当前件复检计数 [次] / the current part recheck count
    nDegradeCnt  : UDINT := 0;  // 累计降级计数 [次] / the accumulated degrade count
    eState       : E_DL_VrgPhase := E_DL_VrgPhase.eVrgIdle; // 流程状态输出 [-] / the process state outlet
    bFault       : BOOL := FALSE; // 故障锁存指示（解除 = bReset 沿）[-] / the fault latch indicator
    bError       : BOOL := FALSE; // 组态域闸故障锁存 [-] / the config gate fault latch
END_VAR
VAR CONSTANT
    DL_VRG_CNTMAX : UDINT := 4294967294; // 计数防回绕上界 [次] / the counter anti wrap clamp bound
END_VAR
VAR
    _ePhase    : E_DL_VrgPhase := E_DL_VrgPhase.eVrgIdle; // 内部相位，CASE 唯一写入目标 / the internal phase, the single CASE write target
    _nRecheck  : INT := 0;   // 复检计数寄存 [次] / the recheck count register
    _bInit     : BOOL := FALSE; // 首拍初始化标志（R310，真实使用：首拍安全态预置）/ the first scan flag, real use
    rtPart     : R_TRIG;     // 到位沿，段 0 无条件刷新 / the part edge
    rtReady    : R_TRIG;     // 结果选通沿，段 0 无条件刷新 / the strobe edge
    rtReset    : R_TRIG;     // 复位沿，段 0 无条件刷新 / the reset edge
    tonJudge   : TON;        // 判决窗，段 0 无条件刷新 / the judge window
END_VAR

// 段 0｜定时器与沿检测无条件周期刷新（禁入分支，R7）/ segment 0, the unconditional refresh
rtPart(CLK := bPartIn); // 到位沿 / the part edge
rtReady(CLK := bResultReady); // 选通沿 / the strobe edge
rtReset(CLK := bReset); // 复位沿 / the reset edge
tonJudge(IN := (_ePhase = E_DL_VrgPhase.eVrgJudge) OR (_ePhase = E_DL_VrgPhase.eVrgRecheck), PT := tJudgeWin); // 判决窗（复检共用不重启，边界二）/ the judge window shared by the recheck

// 段 1｜首拍初始化（R310 真实使用路径）：相位安全态显式预置 / segment 1, the first scan init
IF NOT _bInit THEN // 首拍一拍 / the first scan
    _bInit := TRUE; // 置首拍标志 / raise the flag
    _ePhase := E_DL_VrgPhase.eVrgIdle; // 相位显式安全预置 / the explicit safe preset
END_IF

// 段 2｜组态域闸与复位（边界四，解除路径 = bReset 沿，R188）/ segment 2, the config gate and the reset
IF (nRecheckMax < 0) OR (nRecheckMax > 9) THEN // 复检上限越域 / the recheck bound out of domain
    bError := TRUE; // 置域闸锁存 / raise the config latch
END_IF
IF rtReset.Q THEN // 复位沿 / the reset edge
    bError := FALSE; // 清域闸锁存 / clear the config latch
    _nRecheck := 0; // 清复检计数 / clear the recheck count
    IF _ePhase = E_DL_VrgPhase.eVrgFault THEN // 仅故障相消化复位迁相 / only the fault phase consumes the reset
        _ePhase := E_DL_VrgPhase.eVrgIdle; // 回空闲（解除路径唯一，R188）/ back to idle
    END_IF
END_IF

// 段 3｜单拍脉冲前置清零（边界三，纪律③）/ segment 3, the per scan pulse preset
bPass := FALSE; // 通过脉冲预清零 / preset the pass false
bReject := FALSE; // 拒收脉冲预清零 / preset the reject false
bDegrade := FALSE; // 降级脉冲预清零 / preset the degrade false

// 段 4｜相位机：ENUM + CASE，含 ELSE 非法相位兜底（R6 / R128）/ segment 4, the phase machine
CASE _ePhase OF

E_DL_VrgPhase.eVrgIdle: // 空闲相 / the idle phase
    IF rtPart.Q AND (NOT bError) THEN // 受理到位沿开窗（组态合法）/ accept the part edge
        _nRecheck := 0; // 复检计数清零 / clear the recheck count
        _ePhase := E_DL_VrgPhase.eVrgJudge; // 迁判决窗相 / to the judge phase
    END_IF

E_DL_VrgPhase.eVrgJudge: // 判决窗相 / the judge phase
    IF rtReady.Q THEN // 结果选通 / the result strobe
        IF bVisionOk THEN // 判 OK / the ok verdict
            bPass := TRUE; // 置通过单脉冲 / raise the pass pulse
            _ePhase := E_DL_VrgPhase.eVrgIdle; // 回空闲 / back to idle
        ELSIF _nRecheck < nRecheckMax THEN // NG 且复检额度未用尽 / an NG with the recheck budget left
            _nRecheck := _nRecheck + 1; // 复检计数推进 / advance the recheck count
            _ePhase := E_DL_VrgPhase.eVrgRecheck; // 迁复检窗相（窗续走不重启）/ to the recheck phase
        ELSE // NG 且额度用尽：拒收 / the NG beyond the budget, reject
            bReject := TRUE; // 置拒收单脉冲 / raise the reject pulse
            _ePhase := E_DL_VrgPhase.eVrgIdle; // 回空闲 / back to idle
        END_IF
    ELSIF tonJudge.Q THEN // 窗超时无结果：降级安全侧判 NG（窗口末退出迁移，边界一二）/ the window expired, the safe downgrade
        bDegrade := TRUE; // 置降级单脉冲 / raise the degrade pulse
        bReject := TRUE; // 降级安全侧拒收（R191 降级显式）/ the safe reject
        IF nDegradeCnt < DL_VRG_CNTMAX THEN // 计数防回绕 / the wrap guard
            nDegradeCnt := nDegradeCnt + 1; // 降级计数推进 / advance the degrade count
        END_IF
        _ePhase := E_DL_VrgPhase.eVrgIdle; // 回空闲 / back to idle
    END_IF

E_DL_VrgPhase.eVrgRecheck: // 复检窗相 / the recheck phase
    IF rtReady.Q THEN // 复检结果选通 / the recheck strobe
        IF bVisionOk THEN // 复检判 OK / the recheck ok
            bPass := TRUE; // 置通过单脉冲 / raise the pass pulse
            _ePhase := E_DL_VrgPhase.eVrgIdle; // 回空闲 / back to idle
        ELSE // 复检仍 NG：终判拒收 / the recheck NG, the final reject
            bReject := TRUE; // 置拒收单脉冲 / raise the reject pulse
            _ePhase := E_DL_VrgPhase.eVrgIdle; // 回空闲 / back to idle
        END_IF
    ELSIF tonJudge.Q THEN // 复检窗超时：安全侧拒收（窗口末退出迁移）/ the recheck window expired, the safe reject
        bReject := TRUE; // 置拒收单脉冲 / raise the reject pulse
        _ePhase := E_DL_VrgPhase.eVrgIdle; // 回空闲 / back to idle
    END_IF

E_DL_VrgPhase.eVrgFault: // 故障锁存相：本件无迁入源，保留对称兜底位 / the fault latch phase, reserved symmetric
    // 驻留无动作：迁相由段 2 复位分支消化 / dwell, the migrate in the reset branch

ELSE // 非法相位兜底（R128）/ the illegal phase fallback
    _ePhase := E_DL_VrgPhase.eVrgIdle; // 回空闲安全相 / back to the safe idle
END_CASE

// 段 5｜统一出口（R191 名实双出口）/ segment 5, the unified outlet
nRecheckCnt := _nRecheck; // 复检计数出口 / the recheck count outlet
eState := _ePhase; // 状态出口 / the state outlet
bFault := (_ePhase = E_DL_VrgPhase.eVrgFault); // 故障指示与相位同源 / the fault indicator shares the phase
END_FUNCTION_BLOCK

(* ---- FB_DL_VocVentTrim.st ---- *)
// FB_DL_VocVentTrim v1.0.0
// 开源溯源：self-cleanroom / HVAC 域延伸
(*
  道莅工业代码库 | DL_Process | FB_DL_VocVentTrim
  版本: 1.0.0 | 日期: 2026-11-23 | 轮次: R75
  功能: VOC 浓度需求通风 trim：按 VOC 实测-设定偏差比例调节新风阀开度，
        持续超限升入 boost 相全开，迟滞回落
  邻件关系: 与 RoomCo2DemandVent 同构异介质 —— 差异点：邻件介质为 CO2
            （ppm 域 ~400-2000，比例增益按人体舒适域标定），本件介质为
            VOC（ppb/ppm 域，阈值按工业卫生限值标定，boost 相出口口径
            与换气次数系数独立），控制律同构（比例 trim + 超限 boost），
            码位独立（本件 16#0002_2501，避让 CO2 件码段）
*)
TYPE E_DL_VocVentPhase :
(
    eIdle  := 0,    // 空闲（失能）/ Idle, disabled
    eTrim  := 10,   // 比例 trim 相 / Proportional trim phase
    eBoost := 20,   // 超限 boost 相（全开）/ Boost phase, full open
    eFault := 90    // 故障锁定 / Fault locked
);
END_TYPE

FUNCTION_BLOCK FB_DL_VocVentTrim
VAR_INPUT
    bEnable      : BOOL := FALSE;             // 总使能，FALSE 阀门回最小 / Master enable
    fVocPpm      : REAL := 0.0;               // VOC 实测浓度 [ppm]，域 0..100 / Measured VOC [ppm]
    fVocSetPpm   : REAL := 10.0;              // VOC 设定阈值 [ppm]，域 > 0 / VOC setpoint [ppm]
    fBoostPpm    : REAL := 20.0;              // boost 触发阈值 [ppm]，域 > 设定 / Boost trigger threshold [ppm]
    fTrimGainPct : REAL := 10.0;              // trim 增益 [百分点每 ppm] / Trim gain [pct per ppm]
    fVentMinPct  : REAL := 0.0;               // 新风阀最小开度 [%] / Vent minimum [%]
    fVentMaxPct  : REAL := 100.0;             // 新风阀最大开度 [%] / Vent maximum [%]
    fHystPpm     : REAL := 2.0;               // boost 退出迟滞 [ppm] / Boost exit hysteresis [ppm]
END_VAR
VAR_OUTPUT
    fVentCmdPct  : REAL;                      // 新风阀开度指令 [%] / Vent command [%]
    bBoost       : BOOL;                      // boost 相标志 [-] / Boost phase flag
    bValid       : BOOL;                      // 组态有效回执 [-] / Config validity receipt
    bError       : BOOL;                      // 故障标志，与故障级码配对 / Fault flag paired with fault code
    uErrorId     : UDINT;                     // 事件码，0 = 无事件 / Event code, 0 = none
    eStateOut    : E_DL_VocVentPhase;         // 状态机当前态，段尾单点映射 / Phase mapped at tail
END_VAR
VAR
    _eState      : E_DL_VocVentPhase := E_DL_VocVentPhase.eIdle;   // 内部状态 / Internal state
    bCfgOk       : BOOL;                      // 组态闸结果 [-] / Config gate result
    bMeasOk      : BOOL;                      // 测量域闸结果 [-] / Measurement gate result
    fError       : REAL;                      // 偏差 = 实测 - 设定 [ppm] / Error = measured - setpoint
    fCmd         : REAL;                      // 开度指令暂存 [%] / Command buffer [%]
END_VAR

// —— 段 0：全路径缺省（输出中性值） —— //
fVentCmdPct := fVentMinPct;                   // 开度缺省最小（安全位）/ Command default minimum
bBoost := FALSE;                              // boost 标志预清 / Boost preset
bValid := FALSE;                              // 有效回执预清 / Validity preset
bError := FALSE;                              // 故障预清（组态非法路径置位）/ Fault preset
uErrorId := 16#0000;                          // 事件码预清 / Event code preset

// —— 段 1：组态闸与测量域闸 —— //
bCfgOk := (fVocSetPpm > 0.0) AND (fBoostPpm > fVocSetPpm) AND (fVentMaxPct > fVentMinPct)
          AND (fHystPpm >= 0.0) AND (fVocSetPpm = fVocSetPpm) AND (fBoostPpm = fBoostPpm);   // 组态单调 + NaN 闸 / Config monotonic and NaN gate
bMeasOk := (fVocPpm >= 0.0) AND (fVocPpm <= 100.0) AND (fVocPpm = fVocPpm);   // 测量域闸 / Measurement domain gate
IF NOT bCfgOk THEN
    bValid := FALSE;                          // 组态回执降级 / Validity degraded
    bError := TRUE;                           // 故障级：组态非法 / Fault level: invalid config
    uErrorId := 16#0002_2501;                 // 故障码（25xx 步进）/ Fault code
    fVentCmdPct := fVentMinPct;               // 阀门回最小（安全位）/ Vent to minimum
    RETURN;
END_IF
bValid := TRUE;                               // 组态有效回执 / Validity receipt

// —— 段 2：主状态机（ENUM + CASE，含 ELSE 兜底） —— //
CASE _eState OF
E_DL_VocVentPhase.eIdle :
    fCmd := fVentMinPct;                      // 空闲最小开度（安全位）/ Idle minimum
    IF bEnable AND bMeasOk THEN
        _eState := E_DL_VocVentPhase.eTrim;   // 使能且测量有效进 trim 相 / Enabled with valid measurement
    END_IF

E_DL_VocVentPhase.eTrim :
    IF NOT bMeasOk THEN
        fCmd := fVentMinPct;                  // 测量失效：回安全位（本拍不推进）/ Measurement invalid: safe position
        _eState := E_DL_VocVentPhase.eIdle;   // 回空闲等有效测量（退出条件 1：前置消失）/ Exit condition 1
    ELSIF fVocPpm >= fBoostPpm THEN
        fCmd := fVentMaxPct;                  // 超限：本拍即全开（抢先行为）/ Over limit: full open immediately
        _eState := E_DL_VocVentPhase.eBoost;  // 升入 boost 相 / Enter boost
    ELSE
        fError := fVocPpm - fVocSetPpm;       // 偏差 [ppm] / Error [ppm]
        IF fError < 0.0 THEN
            fError := 0.0;                    // 负偏差不回关（通风只增不减，滞环防抖）/ Nonnegative error
        END_IF
        fCmd := fVentMinPct + fError * fTrimGainPct;   // 比例 trim 指令 / Proportional trim command
        IF fCmd > fVentMaxPct THEN
            fCmd := fVentMaxPct;              // 上限钳位 / Clamp high
        END_IF
        IF fCmd < fVentMinPct THEN
            fCmd := fVentMinPct;              // 下限钳位 / Clamp low
        END_IF
        IF NOT bEnable THEN
            _eState := E_DL_VocVentPhase.eIdle;   // 失能回空闲（退出条件 2）/ Exit condition 2
        END_IF
    END_IF

E_DL_VocVentPhase.eBoost :
    fCmd := fVentMaxPct;                      // boost 相全开 / Boost full open
    bBoost := TRUE;                           // boost 标志 / Boost flag
    IF (NOT bMeasOk) OR (NOT bEnable) THEN
        bBoost := FALSE;                      // 失效/失能退出 boost（退出条件 1）/ Exit on invalid or disabled
        _eState := E_DL_VocVentPhase.eIdle;   // 回空闲 / To idle
    ELSIF fVocPpm < (fBoostPpm - fHystPpm) THEN
        bBoost := FALSE;                      // 浓度低于阈值减迟滞退出（退出条件 2）/ Exit below threshold with hysteresis
        _eState := E_DL_VocVentPhase.eTrim;   // 回 trim 相 / Back to trim
    END_IF

E_DL_VocVentPhase.eFault :
    fCmd := fVentMinPct;                      // 故障相安全位 / Fault safe position
    IF bCfgOk THEN
        _eState := E_DL_VocVentPhase.eIdle;   // 组态恢复解锁回空闲（解除路径可达）/ Unlock on valid config
    END_IF

ELSE
    _eState := E_DL_VocVentPhase.eFault;      // 非法状态拦截 / Illegal state interception
    uErrorId := 16#0002_2501;                 // 故障级：相 ID 越界 / Fault level: phase id out of range
    fCmd := fVentMinPct;                      // 安全位 / Safe position
END_CASE

// —— 段 3：输出映射（段尾单点） —— //
IF NOT bEnable THEN
    fCmd := fVentMinPct;                      // 失能最高优先回安全位 / Disabled highest priority
END_IF
fVentCmdPct := fCmd;                          // 开度指令输出 / Command output
eStateOut := _eState;                         // 输出枚举段尾单点映射 / Tail single-point mapping
END_FUNCTION_BLOCK

(* ---- FB_DL_WaferBreakDetect.st ---- *)
(*
  FB_DL_WaferBreakDetect  —  电池片隐裂/碎片在线判据 / Wafer crack-break online detection
  分类 Category : DL_Process
  码位 Code     : 16#06_0_BB
  段位说明      : R38 W7 预留 B6~BF 本轮正式启用，BA 格由 TankLevelStrapping 启用，本件启用 BB 格
  版本 Version  : 1.0.0
  来源 Source   : t2-1-lgf-measurement — 视觉位 + 峰值捕获双判据聚合分级待挖项
  溯源 Origin   : clean-room 实现，未复制任何源码行
  功能 Function : 1) 视觉结果位判据：FC_DL_BitFieldExtract 从视觉结果字提取碎片位/隐裂位
                  （每片在位沿采样一次，单件瞬时判定）；
                  2) 突发峰值判据：FB_DL_PeakDetector 捕获贴合力信号突发峰值
                  （fPeakThreshN 阈值事件），批内突发异常口径；
                  3) 双判据聚合分级（批内累计口径，非单件越限）：
                  eOk / eWatch / eSuspect / eReject 四级，分级每拍重算；
                  4) 批次管理：bBatchStart 沿清累计，达 uBatchSize 置 bBatchDone。
  边界 Boundary : ① 判据取「批内突发异常」：单件碎片只计件数，分级看批内率，禁单件直接判级；
                  ② 位偏移域闸 0..31（DWORD 字长）；峰值阈值/批量域非法判组态错锁存；
                  ③ 力信号非有限：峰值件内部保持上次有效值（件内防御），本件置信息级码；
                  ④ 无状态机相（聚合型 FB）：分级 CASE 为计算型分类，含 ELSE 兜底；
                  ⑤ R228-B 达标声明：eFault 迁出 = rtReset.Q（输入引脚，恒可达），逐字写于此。
  依赖 Depends  : FC_DL_BitFieldExtract（函数调用，引脚按 registry 实名）；
                  FB_DL_PeakDetector / FB_DL_SignalStatistics（实例化，引脚按 registry 实名）
  码表 Error codes（本件格 06_0_BB，子码步进 +0x100）:
    16#0006_01BB 信息级：批次完成（bBatchDone 置位拍）
    16#0006_02BB 故障级：组态非法（位偏移/阈值/批量域非法），锁存至复位
    16#0006_03BB 信息级：批次分级为拒收（eReject 拍）
    16#0006_04BB 信息级：当前片碎片判定命中
    16#0006_05BB 信息级：突发峰值捕获（批内异常事件）
    16#0006_06BB 信息级：当前片隐裂判定命中
    16#0006_07BB 故障级：保留码，本件无 CASE 主状态机，仅作后续维护者新增分支时的防御式默认码
    16#0006_08BB 故障级：状态机落 ELSE 兜底（分级 CASE 非法分支，防御口径）

  修订历史 Revision :
    2026-11-19  v1.0.0  R39 首版（批次 4 · 序号 19）
*)

TYPE E_DL_WaferGrade :
(
    eOk      := 0,    // 正常：批内无异常累计 / OK, no batch anomalies
    eWatch   := 10,   // 关注：峰值接近阈值（0.8 倍口径）/ Watch, peak near threshold
    eSuspect := 20,   // 可疑：批内有碎片/隐裂/突发累计 / Suspect, batch anomalies present
    eReject  := 30    // 拒收：碎片或突发计数达上限 / Reject, break or burst count at limit
);
END_TYPE

FUNCTION_BLOCK FB_DL_WaferBreakDetect
VAR_INPUT
    uVisionWord   : DWORD := 16#0;      // 视觉结果字（位打包）/ Vision result word, bit-packed
    nBreakBitOff  : INT  := 4;          // 碎片位偏移 [bit]，域 0..31 / Break bit offset
    nCrackBitOff  : INT  := 5;          // 隐裂位偏移 [bit]，域 0..31 / Crack bit offset
    fForceN       : REAL := 0.0;        // 贴合力信号 [N]（突发峰值判据源）/ Lamination force signal
    fPeakThreshN  : REAL := 20.0;       // 突发峰值阈值 [N]，域 > 0 / Burst peak threshold
    bWaferPresent : BOOL := FALSE;      // 当前片在位脉冲（每片一沿）[-] / Wafer present pulse, one edge per piece
    bBatchStart   : BOOL := FALSE;      // 批次启动沿（清批内累计）[-] / Batch start edge, clears batch counters
    uBatchSize    : UDINT := 1000;      // 批量 [片]，域 > 0 / Batch size
    uBreakCntMax  : UDINT := 3;         // 碎片拒收上限 [片]，域 > 0 / Break reject limit
    uBurstCntMax  : UDINT := 5;         // 突发拒收上限 [次]，域 > 0 / Burst reject limit
    bReset        : BOOL := FALSE;      // 故障复位，上升沿生效 / Fault reset, rising edge
END_VAR
VAR_OUTPUT
    bWaferBreak  : BOOL;                // 当前片碎片判定（在位沿采样）[-] / Current-piece break verdict
    bWaferCrack  : BOOL;                // 当前片隐裂判定 [-] / Current-piece crack verdict
    bBurstEvt    : BOOL;                // 突发峰值事件（电平，峰值超阈期间）[-] / Burst event, level while over threshold
    eGrade       : E_DL_WaferGrade;     // 批内分级出口（每拍重算）/ Batch grade outlet, recomputed each scan
    uBreakCnt    : UDINT;               // 批内碎片累计 [片] / Batch break count
    uCrackCnt    : UDINT;               // 批内隐裂累计 [片] / Batch crack count
    uBurstCnt    : UDINT;               // 批内突发累计 [次] / Batch burst count
    uPieceCnt    : UDINT;               // 批内已检片数 [片] / Pieces inspected in batch
    fPeakForceN  : REAL;                // 当前峰值保持值 [N]（峰值件出口）/ Current held peak force
    bBatchDone   : BOOL;                // 批次完成（达批量）[-] / Batch done flag
    bError       : BOOL;                // 故障锁存，仅故障级码置位，bReset 清除 [-] / Fault latch
    uErrorId     : UDINT;               // 事件码，0 = 无事件（故障级锁存回放）/ Event code
END_VAR
VAR
    fbPeak      : FB_DL_PeakDetector;   // 突发峰值捕获实例（主体首部无条件刷新）/ Burst peak detector instance
    fbStat      : FB_DL_SignalStatistics;   // 力信号统计窗实例（主体首部无条件刷新）/ Force statistics window instance
    rtWafer     : R_TRIG;               // 在位脉冲上升沿 / Wafer present rising edge
    rtBatch     : R_TRIG;               // 批次启动上升沿 / Batch start rising edge
    rtReset     : R_TRIG;               // 故障复位上升沿 / Fault reset rising edge
    _uFieldBrk  : DWORD;                // 碎片位提取结果 / Break bit extraction result
    _uMaskBrk   : DWORD;                // 碎片位掩码（件出口）/ Break bit mask
    _nActWBrk   : INT;                  // 碎片位实际宽度 / Break bit actual width
    _uErrBrk    : UDINT;                // 碎片位提取错误码 / Break extraction error
    _bValBrk    : BOOL;                 // 碎片位提取有效 / Break extraction valid
    _uFieldCrk  : DWORD;                // 隐裂位提取结果 / Crack bit extraction result
    _uMaskCrk   : DWORD;                // 隐裂位掩码 / Crack bit mask
    _nActWCrk   : INT;                  // 隐裂位实际宽度 / Crack bit actual width
    _uErrCrk    : UDINT;                // 隐裂位提取错误码 / Crack extraction error
    _bValCrk    : BOOL;                 // 隐裂位提取有效 / Crack extraction valid
    _bBurstLatch: BOOL;                 // 当前片突发锁存（片内保持，沿采样时消费）/ Per-piece burst latch
    _eGradeInt  : E_DL_WaferGrade := E_DL_WaferGrade.eOk;   // 分级内部量（CASE 唯一写入目标）/ Internal grade, sole CASE target
    _uInfo      : UDINT;                // 信息码，每拍重算 / Info code
    _uFault     : UDINT;                // 故障码锁存寄存 / Latched fault code register
    _bFault     : BOOL;                 // 故障锁存位 / Latched fault bit
    _bCfgBad    : BOOL;                 // 组态非法聚合 / Configuration invalid aggregate
END_VAR
VAR CONSTANT
    DL_WBD_INF_CAP   : REAL := 1.0E15;     // 非有限值筛查幅值上限 / Non-finite screening cap
    DL_WBD_BIT_MAX   : INT  := 31;         // 位偏移上限 [bit]（DWORD 字长）/ Bit offset upper bound
    DL_WBD_CNT_MAX   : UDINT := 16#FFFF_FFFE;  // 计数饱和上限 / Counter saturation bound
    DL_WBD_WATCH_RAT : REAL := 0.8;        // 关注级阈值比（峰值/阈值）[无量纲] / Watch-grade threshold ratio
END_VAR

(* —— 段 0：边沿与依赖件实例无条件周期刷新（R182：调用语句不得置于 IF/CASE 内） —— *)
rtWafer(CLK := bWaferPresent);                          // 在位沿刷新，每拍必调
rtBatch(CLK := bBatchStart);                            // 批次沿刷新，每拍必调
rtReset(CLK := bReset);                                 // 复位沿刷新，每拍必调
fbPeak(bEnable := TRUE,                                 // 峰值捕获恒使能
       bReset := rtWafer.Q,                             // 每片在位沿复位峰值（片口径）
       fSignal := fForceN,                              // 贴合力信号
       tSample := T#10MS,                               // 采样周期（标准口径）
       fDecayRate := 0.0,                               // 不衰减（片内保持口径）
       bDetectValley := FALSE,                          // 只测峰
       fThreshold := MAX(fPeakThreshN, 1.0E-6),         // 突发阈值（下限防零阈常报）
       bThresholdEnable := TRUE);                       // 阈值事件使能
fbStat(fIn := fForceN,                                  // 力信号统计窗（诊断随行）
       bSample := TRUE,                                 // 每拍采样
       nWindow := 32,                                   // 窗长（标准口径）
       bClear := rtBatch.Q);                            // 批次沿清窗

(* —— 段 1：单拍量预清零（锁存量 _uFault/_bFault/_uBreakCntInt 等累计量不入清单，R187①） —— *)
_uInfo := 16#0000_0000;             // 信息码每拍重算
_bCfgBad := FALSE;                  // 组态非法预清零
bWaferBreak := FALSE;               // 当前片判定缺省 FALSE（沿采样段单点置位）
bWaferCrack := FALSE;               // 当前片判定缺省 FALSE
bBatchDone := FALSE;                // 批完成缺省 FALSE（计数段单点置位）
uErrorId := 16#0000_0000;           // 事件码缺省无事件

(* —— 段 2：组态域闸（覆盖全部参与判据换算的引脚，R151） —— *)
IF (nBreakBitOff < 0) OR (nBreakBitOff > DL_WBD_BIT_MAX)
   OR (nCrackBitOff < 0) OR (nCrackBitOff > DL_WBD_BIT_MAX) THEN
    _bCfgBad := TRUE;               // 位偏移域非法
END_IF
IF (fPeakThreshN <= 0.0) OR (ABS(fPeakThreshN) > DL_WBD_INF_CAP)
   OR (fForceN <> fForceN) OR (ABS(fForceN) > DL_WBD_INF_CAP) OR ((fForceN - fForceN) <> 0.0) THEN
    _bCfgBad := TRUE;               // 阈值/力信号域非法
END_IF
IF (uBatchSize = 0) OR (uBreakCntMax = 0) OR (uBurstCntMax = 0) THEN
    _bCfgBad := TRUE;               // 批量/上限域非法
END_IF

(* —— 段 3：故障锁存与迁出沿（R228-B：rtReset.Q 恒可达） —— *)
IF _bCfgBad AND (NOT _bFault) THEN
    _uFault := 16#0006_02BB;        // 故障级：组态非法（仅首次进入时写入）
    _bFault := TRUE;
END_IF
IF rtReset.Q AND (NOT _bCfgBad) THEN
    _bFault := FALSE;               // 清故障锁存位（组态恢复合法为前提）
    _uFault := 16#0000_0000;
END_IF

(* —— 段 4：批次启动沿（清批内累计） —— *)
IF rtBatch.Q THEN
    uBreakCnt := 0;                 // 碎片累计清零
    uCrackCnt := 0;                 // 隐裂累计清零
    uBurstCnt := 0;                 // 突发累计清零
    uPieceCnt := 0;                 // 片数清零
    bBatchDone := FALSE;            // 批完成标志复位（沿拍清除）
END_IF

(* —— 段 5：突发峰值判据（峰值件出口镜像 + 批内突发锁存） —— *)
fPeakForceN := fbPeak.fPeak;        // 峰值保持值镜像
bBurstEvt := fbPeak.bOverThreshold; // 超阈电平镜像（每拍重算）
IF bBurstEvt AND (NOT _bBurstLatch) THEN
    _bBurstLatch := TRUE;           // 片内突发锁存（防同一突发重复计数）
    uBurstCnt := uBurstCnt + 1;     // 批内突发累计
    IF uBurstCnt >= DL_WBD_CNT_MAX THEN
        uBurstCnt := DL_WBD_CNT_MAX;    // 计数饱和防回绕
    END_IF
    _uInfo := 16#0006_05BB;         // 信息级：突发峰值捕获
END_IF
IF rtWafer.Q THEN
    _bBurstLatch := FALSE;          // 片沿：突发锁存复位（下一片重新捕获）
END_IF

(* —— 段 6：视觉位判据（在位沿采样一次；位段提取原子 ×2） —— *)
IF rtWafer.Q AND (NOT _bFault) THEN
    FC_DL_BitFieldExtract(uSource := uVisionWord,       // 视觉结果字
                          nOffset := nBreakBitOff,      // 碎片位偏移
                          nWidth := 1,                  // 单位提取
                          uField => _uFieldBrk,         // 提取结果
                          uMask => _uMaskBrk,           // 掩码
                          nActualW => _nActWBrk,        // 实际宽度
                          uErrorId => _uErrBrk,         // 错误码
                          bValid => _bValBrk);          // 有效标志
    FC_DL_BitFieldExtract(uSource := uVisionWord,       // 视觉结果字
                          nOffset := nCrackBitOff,      // 隐裂位偏移
                          nWidth := 1,                  // 单位提取
                          uField => _uFieldCrk,         // 提取结果
                          uMask => _uMaskCrk,           // 掩码
                          nActualW => _nActWCrk,        // 实际宽度
                          uErrorId => _uErrCrk,         // 错误码
                          bValid => _bValCrk);          // 有效标志
    IF _bValBrk AND (_uFieldBrk > 0) THEN
        bWaferBreak := TRUE;        // 当前片碎片判定命中
        uBreakCnt := uBreakCnt + 1; // 批内碎片累计
        IF uBreakCnt >= DL_WBD_CNT_MAX THEN
            uBreakCnt := DL_WBD_CNT_MAX;
        END_IF
        _uInfo := 16#0006_04BB;     // 信息级：碎片命中
    END_IF
    IF _bValCrk AND (_uFieldCrk > 0) THEN
        bWaferCrack := TRUE;        // 当前片隐裂判定命中
        uCrackCnt := uCrackCnt + 1; // 批内隐裂累计
        IF uCrackCnt >= DL_WBD_CNT_MAX THEN
            uCrackCnt := DL_WBD_CNT_MAX;
        END_IF
        _uInfo := 16#0006_06BB;     // 信息级：隐裂命中
    END_IF
    uPieceCnt := uPieceCnt + 1;     // 已检片数
    IF uPieceCnt >= DL_WBD_CNT_MAX THEN
        uPieceCnt := DL_WBD_CNT_MAX;
    END_IF
END_IF

(* —— 段 7：分级 CASE（计算型分类，含 ELSE 兜底） —— *)
IF (NOT _bFault) AND (uPieceCnt > 0) THEN
    CASE _eGradeInt OF
    E_DL_WaferGrade.eOk:
        IF (uBreakCnt >= uBreakCntMax) OR (uBurstCnt >= uBurstCntMax) THEN
            _eGradeInt := E_DL_WaferGrade.eReject;      // 达拒收上限：进拒收级
        ELSIF (uBreakCnt > 0) OR (uCrackCnt > 0) OR (uBurstCnt > 0) THEN
            _eGradeInt := E_DL_WaferGrade.eSuspect;     // 有异常累计：进可疑级
        ELSIF fPeakForceN >= fPeakThreshN * DL_WBD_WATCH_RAT THEN
            _eGradeInt := E_DL_WaferGrade.eWatch;       // 峰值近阈：进关注级
        END_IF
    E_DL_WaferGrade.eWatch:
        IF (uBreakCnt >= uBreakCntMax) OR (uBurstCnt >= uBurstCntMax) THEN
            _eGradeInt := E_DL_WaferGrade.eReject;      // 达拒收上限：进拒收级
        ELSIF (uBreakCnt > 0) OR (uCrackCnt > 0) OR (uBurstCnt > 0) THEN
            _eGradeInt := E_DL_WaferGrade.eSuspect;     // 有异常累计：进可疑级
        ELSIF fPeakForceN < fPeakThreshN * DL_WBD_WATCH_RAT THEN
            _eGradeInt := E_DL_WaferGrade.eOk;          // 峰值回落：回正常级
        END_IF
    E_DL_WaferGrade.eSuspect:
        IF (uBreakCnt >= uBreakCntMax) OR (uBurstCnt >= uBurstCntMax) THEN
            _eGradeInt := E_DL_WaferGrade.eReject;      // 达拒收上限：进拒收级
        END_IF
    E_DL_WaferGrade.eReject:
        IF rtBatch.Q THEN
            _eGradeInt := E_DL_WaferGrade.eOk;          // 新批次：回正常级（段 4 清累计后自然满足）
        END_IF
    ELSE
        _uFault := 16#0006_08BB;    // 故障级：非法分级 ID 兜底
        _bFault := TRUE;
        _eGradeInt := E_DL_WaferGrade.eReject;      // 防御口径：回拒收级
    END_CASE
    IF _eGradeInt = E_DL_WaferGrade.eReject THEN
        _uInfo := 16#0006_03BB;     // 信息级：分级拒收（覆盖命中码，分级状态优先）
    END_IF
END_IF

(* —— 段 8：批次完成（达批量置位，新批次沿清除） —— *)
IF (NOT _bFault) AND (uPieceCnt >= uBatchSize) THEN
    bBatchDone := TRUE;             // 批完成标志
    _uInfo := 16#0006_01BB;         // 信息级：批次完成（覆盖分级码，完成事件优先）
END_IF

(* —— 段 9：出口单点映射（名实同源；锁存码回放，禁同拍抹除） —— *)
eGrade := _eGradeInt;               // 分级出口镜像
IF _bFault THEN
    uErrorId := _uFault;            // 故障锁存码回放
    bError := TRUE;
    bBatchDone := FALSE;            // 故障态批完成强制 FALSE（安全侧）
ELSE
    uErrorId := _uInfo;             // 信息码
    bError := FALSE;
END_IF

END_FUNCTION_BLOCK

(* ---- FB_DL_WaferCountPreset.st ---- *)
(*
  FB_DL_WaferCountPreset  —  晶圆计数预置饱和（预置计满 + 花篮位模计数） / Wafer preset count with saturation and cassette-slot modulo counting
  分类 Category : DL_Process
  版本 Version  : 1.0.0
  来源 Source   : t2-1-lgf-counter — 计数族深化（与 WaferCountAxis/WaferCountYield 分工：那两件管计数轴/良率统计，本件管预置饱和与模计数）
  溯源 Origin   : clean-room 实现，未复制任何源码行
  功能 Function : 1) 预置计数：bCntPulse 上升沿递增 uCount，达 uPreset 置 bPresetDone
                  并停计；计满后仍来沿 → 0380 溢出饱和锁存（防静默丢片）；
                  2) 花篮位模计数：bSlotPulse 沿按 uCassSlots 取模递增 uCassMod，
                  回零拍发信息级 04A8；模基数域闸 uCassSlots > 0；
                  3) 脉冲宽度监视：计数沿后高电平持续超 tMinPulse → 0381 锁存
                  （同拍重触发漏计风险，归因独立）；
                  4) 相位机：eIdle → eCount → eFull → eFault；
                  5) 解除式全当拍量（R240 落地），逐 BOOL 标注见段 4。
  边界 Boundary : ① 组态闸：uPreset = 0 或 uCassSlots = 0 或 tMinPulse <= 0
                  → 037F 锁存，ELSE 兜底归并 037F（码表声明）；
                  ② 模计数用 MOD 内建，模基数 > 0 已由域闸保证，无除零路径；
                  ③ 计数沿 R_TRIG 与宽度监视 TON 均无条件周期刷新；
                  ④ 无 GVL 依赖：纯引脚输入输出，无外部变量引用，无物理 IO 地址。
  依赖 Depends  : Standard.library（TON / R_TRIG）
  码表 Error codes（Process 段 0005，窗口 037F~0381 / 04A7~04A9）:
    16#0005_037F 故障级：组态非法（预置/模基数/最小脉宽域非法）或相位落 ELSE 兜底（归并声明），锁存至 bReset
    16#0005_0380 故障级：预置计满后计数沿溢出锁存，锁存至 bReset
    16#0005_0381 故障级：计数脉冲宽度异常锁存（高电平持续超 tMinPulse），锁存至 bReset
    16#0005_04A7 信息级：预置计满沿（进 eFull）
    16#0005_04A8 信息级：花篮模计数回零沿
    16#0005_04A9 信息级：计数复位完成沿
  修订历史 Revision :
    2026-11-19  v1.0.0  R42 首版（批次 2 · 序号 1）
*)

TYPE E_DL_WcpState :
(
    eIdle   := 0,    // 未使能：不计数 / Idle, not counting
    eCount  := 10,   // 计数中：沿递增 / Counting, edge increments
    eFull   := 20,   // 计满：预置达成停计 / Full, preset reached
    eFault  := 90    // 故障：溢出或脉宽锁定 / Fault, latched
);
END_TYPE

FUNCTION_BLOCK FB_DL_WaferCountPreset
VAR_INPUT
    bCntPulse    : BOOL := FALSE;     // 晶圆计数脉冲 [-] / Wafer count pulse
    bSlotPulse   : BOOL := FALSE;     // 花篮槽位脉冲 [-] / Cassette slot pulse
    uPreset      : UDINT := 25;       // 预置计数值 [片]，域 > 0 / Preset count value
    uCassSlots   : UDINT := 25;       // 花篮模计数基数 [槽]，域 > 0 / Cassette modulo base
    tMinPulse    : TIME := T#5MS;     // 最小合法脉宽 [ms]，域 > 0 / Minimum legal pulse width
    bCntEn       : BOOL := FALSE;     // 计数使能（电平）[-] / Count enable, level
    bCntRst      : BOOL := FALSE;     // 计数复位指令，上升沿清计数 [-] / Count reset command edge
    bReset       : BOOL := FALSE;     // 复位，上升沿清故障锁存 / Reset edge clears fault latch
END_VAR
VAR_OUTPUT
    eState       : E_DL_WcpState;     // 状态出口，段尾单点映射 / State outlet
    uCount       : UDINT;             // 晶圆计数 [片] / Wafer count
    bPresetDone  : BOOL;              // 预置达成标志（eFull 相电平）[-] / Preset-done flag
    uCassMod     : UDINT;             // 花篮模计数值 [槽] / Cassette modulo count
    bError       : BOOL;              // 故障锁存标志 / Fault latch flag
    nErrId       : UDINT;             // 事件码，0 = 无事件 / Event code
END_VAR
VAR
    tonPulseW    : TON;               // 脉冲宽度监视（电平式），无条件刷新 / Pulse width watch timer
    rtCntPulse   : R_TRIG;            // 计数脉冲沿实例，无条件刷新 / Count pulse edge instance
    rtSlotPulse  : R_TRIG;            // 槽位脉冲沿实例，无条件刷新 / Slot pulse edge instance
    rtCntRst     : R_TRIG;            // 计数复位沿实例，无条件刷新 / Count reset edge instance
    rtReset      : R_TRIG;            // 复位沿实例，无条件刷新 / Reset edge instance
    _eState      : E_DL_WcpState := E_DL_WcpState.eIdle;  // 内部相位（CASE 唯一写入目标）/ Internal phase
    _bFault      : BOOL;              // 故障锁存位（锁存量）/ Latched fault bit
    _uFault      : UDINT;             // 故障码锁存（锁存量）/ Latched fault code
    _uInfo       : UDINT;             // 信息码，每拍重算 / Transient info code
END_VAR

(* —— 段 0：定时器与沿实例无条件周期刷新（禁置于 IF/CASE 内） —— *)
rtCntPulse(CLK := bCntPulse);                            // 计数脉冲沿（每拍必调）
rtSlotPulse(CLK := bSlotPulse);                          // 槽位脉冲沿（每拍必调）
rtCntRst(CLK := bCntRst);                                // 计数复位沿（每拍必调）
rtReset(CLK := bReset);                                  // 复位沿（每拍必调）
tonPulseW(IN := bCntPulse, PT := tMinPulse);             // 脉宽监视（电平式，脉冲撤销自动断 IN）

(* —— 段 1：单拍量预清零（锁存量 _bFault/_uFault 不入清单，禁同拍抹除） —— *)
_uInfo := 16#0000_0000;             // 信息码每拍重算
bPresetDone := FALSE;               // 预置达成标志缺省 FALSE
nErrId := 16#0000_0000;             // 事件码缺省无事件

(* —— 段 2：复位沿 + 组态域闸 + 计数复位（判据当拍量） —— *)
IF rtReset.Q THEN                   // rtReset.Q = 当拍量
    _bFault := FALSE;               // 清故障锁存位
    _uFault := 16#0000_0000;        // 清故障锁存码
END_IF
IF (uPreset = 0) OR (uCassSlots = 0) OR (TIME_TO_DINT(tMinPulse) <= 0) THEN
    _uFault := 16#0005_037F;        // 故障级：组态非法
    _bFault := TRUE;                // 故障标志与码位配对（R45）
END_IF
IF rtCntRst.Q THEN                  // 计数复位沿（当拍量）
    uCount := 16#0000_0000;         // 计数清零
    uCassMod := 16#0000_0000;       // 模计数清零
    _uInfo := 16#0005_04A9;         // 信息级：计数复位完成沿
END_IF

(* —— 段 3：溢出与脉宽锁存（判据当拍量/电平式窗） —— *)
IF (NOT _bFault) AND tonPulseW.Q THEN
    _uFault := 16#0005_0381;        // 故障级：脉宽异常（同拍重触发漏计风险）
    _bFault := TRUE;
END_IF
IF (NOT _bFault) AND (_eState = E_DL_WcpState.eFull) AND rtCntPulse.Q THEN
    _uFault := 16#0005_0380;        // 故障级：计满后计数沿溢出
    _bFault := TRUE;
END_IF

(* —— 段 4：故障解除式（R240 落地，逐 BOOL 标注）：
     rtReset.Q = 当拍量；NOT bCntPulse = 当拍量；NOT bCntEn = 当拍量。
     均不含锁存量（_bFault/_uFault），解除边真实可达（脉冲撤销 + 撤使能 + 复位沿）。 —— *)
IF rtReset.Q AND (NOT bCntPulse) AND (NOT bCntEn) THEN
    _bFault := FALSE;               // 清故障锁存位（锁存量，仅此当拍量解除沿可清）
    _uFault := 16#0000_0000;        // 清故障锁存码（锁存量，仅本当拍量解除沿可清）
    IF _eState = E_DL_WcpState.eFault THEN
        _eState := E_DL_WcpState.eIdle;     // 故障相迁出：回未使能
    END_IF
END_IF

(* —— 段 5：相位机（CASE 全覆盖 + ELSE 兜底） —— *)
CASE _eState OF

E_DL_WcpState.eIdle:
    IF bCntEn AND (NOT _bFault) THEN
        _eState := E_DL_WcpState.eCount;    // 使能：进计数相
    END_IF

E_DL_WcpState.eCount:
    IF rtCntPulse.Q THEN                    // 计数沿（当拍量）
        IF uCount < uPreset THEN
            uCount := uCount + 1;           // 计数递增（先比后加，防跨预置）
        END_IF
        IF uCount >= uPreset THEN
            _uInfo := 16#0005_04A7;         // 信息级：预置计满沿
            _eState := E_DL_WcpState.eFull; // 进计满相
        END_IF
    END_IF

E_DL_WcpState.eFull:
    bPresetDone := TRUE;                    // 预置达成标志（相电平）
    IF rtCntPulse.Q THEN
        _uFault := 16#0005_0380;            // 故障级：计满后溢出（段 3 同判据冗余收敛，单点归因）
        _bFault := TRUE;
    END_IF
    IF NOT bCntEn THEN
        _eState := E_DL_WcpState.eIdle;     // 撤使能：回未使能相
    END_IF

E_DL_WcpState.eFault:
    ;                                       // 故障相：等解除沿（段 4 承载迁出）

ELSE
    _uFault := 16#0005_037F;                // 故障级：非法相位兜底（归并组态码，码表声明）
    _bFault := TRUE;
    _eState := E_DL_WcpState.eFault;        // 强制回故障相

END_CASE

(* —— 段 5b：花篮模计数（独立于相位机；模回零沿当拍检出） —— *)
IF (_eState = E_DL_WcpState.eCount) AND rtSlotPulse.Q THEN
    uCassMod := (uCassMod + 1) MOD uCassSlots;  // 模计数（模基数域闸 > 0，无除零）
    IF uCassMod = 0 THEN                        // 回零拍（模运算整型判等合规）
        _uInfo := 16#0005_04A8;                 // 信息级：花篮模回零沿
    END_IF
END_IF

(* —— 段 6：出口单点映射（名实同源；锁存码回放，禁同拍抹除） —— *)
IF _bFault THEN
    nErrId := _uFault;              // 故障锁存码回放
    bPresetDone := FALSE;           // 故障相预置达成出口强制 FALSE（安全侧）
ELSE
    nErrId := _uInfo;               // 信息码
END_IF
bError := _bFault;                  // 故障标志与锁存位同源
eState := _eState;                  // 状态出口单点映射

END_FUNCTION_BLOCK

(* ---- FB_DL_WaferScanRouter.st ---- *)
// =====================================================================
// FB_DL_WaferScanRouter.st
// 晶圆盒扫码路由（扫码契约 + 花篮位取模索引 + 分道路由）
// Wafer cassette scan routing with modulo slot index
// 所属子库: DL_Process    版本: v1.0.0    兼容: CODESYS V3.5+ / TwinCAT 3 / 汇川 InoProShop
// 码位: 16#0005_0467 ~ 16#0005_046B (本件独占 5 槽, 勿复用)
// 溯源: 道莅 clean-room 防御性实现
//       来源组标签: semiconductor, barcode-routing, modulo-index, wafer
// 修改记录: R30 初版 (ROUND_PLAN_R30 序 6)
// =====================================================================
FUNCTION_BLOCK FB_DL_WaferScanRouter
VAR_INPUT
    bScanTrigger : BOOL  := FALSE;  // 扫码触发沿 / Scan trigger edge
    sBarcode     : STRING := '';    // 条码内容（扫码器回读注入）/ Barcode content injected
    bReadOk      : BOOL  := FALSE;  // 读码有效标志 / Read valid flag
    uStationMod  : USINT := 1;      // 花篮位号 1~25, 0 = 组态非法 / Station number 1..25
    abRouteEn    : ARRAY[1..8] OF BOOL;  // 分道允许表, 位序对应分道 1..8 / Route enable table 1..8
    tScanTimeout : TIME  := T#2S;   // 扫码超时窗 T#10MS~T#60S / Scan timeout window [s]
END_VAR
VAR_OUTPUT
    uRouteSel    : USINT := 0;      // 选中分道 1~8, 0 = 拒收 / Selected route, 0 = reject
    bRouteOk     : BOOL  := FALSE;  // 路由成功标志 / Route accepted flag
    uSlotIdx     : USINT := 0;      // 花篮位取模索引 1~8 / Modulo slot index 1..8
    eErr         : UDINT := 16#0005_0467;  // 错误码 / Error code
END_VAR
VAR
    rtrScan      : R_TRIG;          // 扫码触发沿检测, 每拍无条件刷新 / Scan trigger edge, refreshed every cycle
    rtrRead      : R_TRIG;          // 读码有效沿检测, 每拍无条件刷新 / Read-valid edge, refreshed every cycle
    tonScan      : TON;             // 扫码超时定时器, 每拍无条件刷新 / Scan timeout timer, refreshed every cycle
    xBusy        : BOOL  := FALSE;  // 扫码窗进行中标志 / Scan window busy flag
    uRouteCnt    : USINT := 0;      // 使能分道计数 0~8 / Enabled route count 0..8
    uSlotCalc    : USINT := 1;      // 取模索引计算临时量 / Slot index calculation temporary
    uGuard       : USINT := 0;      // 条件减法守卫计数 / Conditional subtraction guard counter
    uZi          : INT   := 1;      // 1..8 数组下标 / Array subscript 1..8
END_VAR

// ---------------------------------------------------------------------
// 代码位表（本件独占, 勿复用）:
//   16#0005_0467 信息 路由成功
//   16#0005_0468 信息 组态非法拒收（花篮位号为 0 或分道全禁用）
//   16#0005_0469 故障 扫码超时未读（拒收）; 码随最近一次判定保持, 重新触发扫码即刷新解除
//   16#0005_046A 信息 读码失败拒收（条码数据在而有效标志为假, 与空串语义分离）
//   16#0005_046B 信息 空条码拒收（读码有效但条码长度为零）
// ---------------------------------------------------------------------

// ---- 分道使能计数 / Enabled route count ----
uRouteCnt := 0;                     // 计数复位 / Reset count
FOR uZi := 1 TO 8 DO
    IF abRouteEn[uZi] THEN
        uRouteCnt := uRouteCnt + 1; // 累计使能分道 / Count enabled route
    END_IF
END_FOR

// ---- 边沿与定时器实例无条件周期刷新（调用不进任何 IF 分支）/ Unconditional edge and timer refresh ----
rtrScan(CLK := bScanTrigger);       // 扫码触发沿 / Scan trigger edge
rtrRead(CLK := bReadOk);            // 读码有效沿 / Read valid edge
tonScan(IN := xBusy, PT := tScanTimeout);   // 扫码窗计时 / Scan window timing

// ---- 触发沿启动扫码窗 / Trigger edge starts scan window ----
IF rtrScan.Q THEN
    xBusy := TRUE;                  // 拍 N 进入扫码窗 / Enter scan window
END_IF

// ---- 扫码窗内判定 / Judgement inside scan window ----
IF xBusy THEN
    IF tonScan.Q THEN
        // 本拍行为: 超时拒收并关窗 / Timeout reject and close window
        uRouteSel := 0;             // 拒收 / Reject
        uSlotIdx  := 0;             // 索引无效 / Index void
        bRouteOk  := FALSE;         // 路由失败 / Route failed
        eErr      := 16#0005_0469;  // 扫码超时 / Scan timeout
        xBusy     := FALSE;         // 拍 N+1 窗关闭, 等下次触发 / Window closed
    ELSIF bReadOk AND (LEN(sBarcode) = 0) THEN
        // 空条码: 读码有效但无内容 / Empty barcode: valid flag but no content
        uRouteSel := 0;
        uSlotIdx  := 0;
        bRouteOk  := FALSE;
        eErr      := 16#0005_046B;  // 空条码拒收 / Empty barcode reject
        xBusy     := FALSE;
    ELSIF (NOT bReadOk) AND (LEN(sBarcode) > 0) THEN
        // 读码失败: 数据在而有效标志为假 / Read failed: data present, valid flag false
        uRouteSel := 0;
        uSlotIdx  := 0;
        bRouteOk  := FALSE;
        eErr      := 16#0005_046A;  // 读码失败拒收 / Read-fail reject
        xBusy     := FALSE;
    ELSIF bReadOk AND (LEN(sBarcode) > 0) THEN
        // 读码成功: 组态校验后路由 / Read ok: config check then route
        IF (uStationMod = 0) OR (uRouteCnt = 0) THEN
            uRouteSel := 0;         // 组态非法拒收 / Config illegal reject
            uSlotIdx  := 0;
            bRouteOk  := FALSE;
            eErr      := 16#0005_0468;
        ELSE
            // 取模索引: 条件减法实现, 不用取余运算（跨平台负数歧义禁令）
            // Modulo by conditional subtraction, no remainder operator
            uSlotCalc := uStationMod;       // 从花篮位号起算 / Start from station number
            uGuard    := 0;                 // 守卫计数清零 / Clear guard
            WHILE (uSlotCalc > uRouteCnt) AND (uGuard < 32) DO
                uSlotCalc := uSlotCalc - uRouteCnt;     // 减一轮分道数 / Subtract one route round
                uGuard    := uGuard + 1;                // 守卫计数防死循环 / Guard against dead loop
            END_WHILE
            uSlotIdx := uSlotCalc;      // 输出取模索引 1..分道数 / Output slot index
            // 路由选择: 升序取首个使能分道 / Route select: first enabled ascending
            uRouteSel := 0;
            FOR uZi := 1 TO 8 DO
                IF (uRouteSel = 0) AND abRouteEn[uZi] THEN
                    uRouteSel := INT_TO_USINT(uZi);     // 首个使能分道 / First enabled route
                END_IF
            END_FOR
            bRouteOk := TRUE;           // 路由成功 / Route accepted
            eErr     := 16#0005_0467;   // 正常码 / Normal code
        END_IF
        xBusy := FALSE;                 // 判定完成关窗 / Judgement done, close window
    END_IF
END_IF

END_FUNCTION_BLOCK
